      W_g[13,36] := 0.38792211;
      W_g[13,37] := -0.01284714;
      W_g[13,38] := -0.07044123;
      W_g[13,39] := -0.01824626;
      W_g[14,0] := 0.11452243;
      W_g[14,1] := -0.08958103;
      W_g[14,2] := 0.00742450;
      W_g[14,3] := -0.03061342;
      W_g[14,4] := 0.01046369;
      W_g[14,5] := -0.11585659;
      W_g[14,6] := -0.20829633;
      W_g[14,7] := -0.23606929;
      W_g[14,8] := 0.00405464;
      W_g[14,9] := -0.14249870;
      W_g[14,10] := 0.44500434;
      W_g[14,11] := -0.01216610;
      W_g[14,12] := 0.02130103;
      W_g[14,13] := 0.01377995;
      W_g[14,14] := -0.06184130;
      W_g[14,15] := -0.00823075;
      W_g[14,16] := -0.01915279;
      W_g[14,17] := -0.04558576;
      W_g[14,18] := 0.06331799;
      W_g[14,19] := 0.08152927;
      W_g[14,20] := 0.53168559;
      W_g[14,21] := 0.26574171;
      W_g[14,22] := -0.16918069;
      W_g[14,23] := -0.07620575;
      W_g[14,24] := 0.06382546;
      W_g[14,25] := 0.06389488;
      W_g[14,26] := -0.00257182;
      W_g[14,27] := -0.51656342;
      W_g[14,28] := -0.13776320;
      W_g[14,29] := -0.24295253;
      W_g[14,30] := -0.07003054;
      W_g[14,31] := -0.24279301;
      W_g[14,32] := -0.02749909;
      W_g[14,33] := 0.02581101;
      W_g[14,34] := -0.14111596;
      W_g[14,35] := 0.25200224;
      W_g[14,36] := 0.05485417;
      W_g[14,37] := 0.20230512;
      W_g[14,38] := 0.05531698;
      W_g[14,39] := 0.08741502;
      W_g[15,0] := 0.09134059;
      W_g[15,1] := 0.23798586;
      W_g[15,2] := -0.21710049;
      W_g[15,3] := 0.01671123;
      W_g[15,4] := -0.06627945;
      W_g[15,5] := 0.03637264;
      W_g[15,6] := -0.06409252;
      W_g[15,7] := 0.00869699;
      W_g[15,8] := 0.06247383;
      W_g[15,9] := 0.02281686;
      W_g[15,10] := -0.03344842;
      W_g[15,11] := 0.25090969;
      W_g[15,12] := 0.23236279;
      W_g[15,13] := -0.16730684;
      W_g[15,14] := 0.02698623;
      W_g[15,15] := -0.12334466;
      W_g[15,16] := -0.08336571;
      W_g[15,17] := 0.02588012;
      W_g[15,18] := 0.18191151;
      W_g[15,19] := -0.02410393;
      W_g[15,20] := -0.01209911;
      W_g[15,21] := 0.03851634;
      W_g[15,22] := 0.03899917;
      W_g[15,23] := -0.03513279;
      W_g[15,24] := -0.00729930;
      W_g[15,25] := -0.10642073;
      W_g[15,26] := -0.05139272;
      W_g[15,27] := -0.04481147;
      W_g[15,28] := 0.00286298;
      W_g[15,29] := 0.04913988;
      W_g[15,30] := 0.03607814;
      W_g[15,31] := -0.06170525;
      W_g[15,32] := -0.01997224;
      W_g[15,33] := -0.01920844;
      W_g[15,34] := -0.18122375;
      W_g[15,35] := -0.04529240;
      W_g[15,36] := -0.02951458;
      W_g[15,37] := -0.04119204;
      W_g[15,38] := 0.24360354;
      W_g[15,39] := -0.01501589;
      W_g[16,0] := 0.03330758;
      W_g[16,1] := 0.03378529;
      W_g[16,2] := -0.01803414;
      W_g[16,3] := 0.07683524;
      W_g[16,4] := -0.00690420;
      W_g[16,5] := 0.06186575;
      W_g[16,6] := -0.05324589;
      W_g[16,7] := 0.00639146;
      W_g[16,8] := -0.03105667;
      W_g[16,9] := -0.02839811;
      W_g[16,10] := -0.02821902;
      W_g[16,11] := 0.34098804;
      W_g[16,12] := 0.27613014;
      W_g[16,13] := 0.05372236;
      W_g[16,14] := -0.07848245;
      W_g[16,15] := 0.19472931;
      W_g[16,16] := 0.02947051;
      W_g[16,17] := 0.30273750;
      W_g[16,18] := -0.21194892;
      W_g[16,19] := -0.39211345;
      W_g[16,20] := 0.05004872;
      W_g[16,21] := -0.00701097;
      W_g[16,22] := -0.05493126;
      W_g[16,23] := -0.06638756;
      W_g[16,24] := 0.04953207;
      W_g[16,25] := -0.07040619;
      W_g[16,26] := 0.02371565;
      W_g[16,27] := 0.05669258;
      W_g[16,28] := 0.01683023;
      W_g[16,29] := 0.01049871;
      W_g[16,30] := -0.03757136;
      W_g[16,31] := -0.14508742;
      W_g[16,32] := 0.06499721;
      W_g[16,33] := 0.04419298;
      W_g[16,34] := 0.17147748;
      W_g[16,35] := 0.11538684;
      W_g[16,36] := -0.02263807;
      W_g[16,37] := 0.09602714;
      W_g[16,38] := -0.19564001;
      W_g[16,39] := -0.07901151;
      W_g[17,0] := -0.29499203;
      W_g[17,1] := -0.13629365;
      W_g[17,2] := 0.12754540;
      W_g[17,3] := -0.06893644;
      W_g[17,4] := 0.12316505;
      W_g[17,5] := -0.05960383;
      W_g[17,6] := 0.20034896;
      W_g[17,7] := -0.04356226;
      W_g[17,8] := 0.02703761;
      W_g[17,9] := 0.06460494;
      W_g[17,10] := 0.13004684;
      W_g[17,11] := 0.24505885;
      W_g[17,12] := -0.04222988;
      W_g[17,13] := -0.06719559;
      W_g[17,14] := -0.02482782;
      W_g[17,15] := 0.21142994;
      W_g[17,16] := -0.06490519;
      W_g[17,17] := -0.00718676;
      W_g[17,18] := -0.06072595;
      W_g[17,19] := 0.09942021;
      W_g[17,20] := 0.12877691;
      W_g[17,21] := -0.55509835;
      W_g[17,22] := 0.01808993;
      W_g[17,23] := -0.10264266;
      W_g[17,24] := -0.39161390;
      W_g[17,25] := -0.18429647;
      W_g[17,26] := 0.28592888;
      W_g[17,27] := 0.28200120;
      W_g[17,28] := -0.28280002;
      W_g[17,29] := 0.37366402;
      W_g[17,30] := -0.26108804;
      W_g[17,31] := -0.16473882;
      W_g[17,32] := -0.02813312;
      W_g[17,33] := 0.06121552;
      W_g[17,34] := -0.13777223;
      W_g[17,35] := 0.06097139;
      W_g[17,36] := -0.11655490;
      W_g[17,37] := 0.32778808;
      W_g[17,38] := -0.00997418;
      W_g[17,39] := 0.61113542;
      W_g[18,0] := -0.28768328;
      W_g[18,1] := 0.04952108;
      W_g[18,2] := 0.27538794;
      W_g[18,3] := 0.13723339;
      W_g[18,4] := -0.17335135;
      W_g[18,5] := 0.00670465;
      W_g[18,6] := 0.08641540;
      W_g[18,7] := -0.07883801;
      W_g[18,8] := 0.03116638;
      W_g[18,9] := -0.13738742;
      W_g[18,10] := 0.04719661;
      W_g[18,11] := -0.16387163;
      W_g[18,12] := 0.33639768;
      W_g[18,13] := 0.00474426;
      W_g[18,14] := 0.00756510;
      W_g[18,15] := 0.14428972;
      W_g[18,16] := -0.27880877;
      W_g[18,17] := 0.02302493;
      W_g[18,18] := -0.08590068;
      W_g[18,19] := -0.09520416;
      W_g[18,20] := -0.04702628;
      W_g[18,21] := -0.21427108;
      W_g[18,22] := -0.01308084;
      W_g[18,23] := -0.13671976;
      W_g[18,24] := -0.33657643;
      W_g[18,25] := -0.29697937;
      W_g[18,26] := -0.38845918;
      W_g[18,27] := -0.13320677;
      W_g[18,28] := 0.12394036;
      W_g[18,29] := -0.01619850;
      W_g[18,30] := -0.00443483;
      W_g[18,31] := 0.02029626;
      W_g[18,32] := -0.14898181;
      W_g[18,33] := -0.13671023;
      W_g[18,34] := -0.39283904;
      W_g[18,35] := -0.18510637;
      W_g[18,36] := 0.02999584;
      W_g[18,37] := -0.09973078;
      W_g[18,38] := -0.00653579;
      W_g[18,39] := 0.00375571;
      W_g[19,0] := -0.11157153;
      W_g[19,1] := 0.03151476;
      W_g[19,2] := -0.09300674;
      W_g[19,3] := -0.03647256;
      W_g[19,4] := 0.28257591;
      W_g[19,5] := 0.03472368;
      W_g[19,6] := -0.19133006;
      W_g[19,7] := 0.01238337;
      W_g[19,8] := 0.10695083;
      W_g[19,9] := 0.06876826;
      W_g[19,10] := -0.15979454;
      W_g[19,11] := 0.04513165;
      W_g[19,12] := -0.09798693;
      W_g[19,13] := 0.24185713;
      W_g[19,14] := -0.15790631;
      W_g[19,15] := -0.06232450;
      W_g[19,16] := -0.01514155;
      W_g[19,17] := -0.04614652;
      W_g[19,18] := -0.04110415;
      W_g[19,19] := -0.02570745;
      W_g[19,20] := 0.10103595;
      W_g[19,21] := -0.08295028;
      W_g[19,22] := 0.07743288;
      W_g[19,23] := -0.15730743;
      W_g[19,24] := 0.17693761;
      W_g[19,25] := 0.33892640;
      W_g[19,26] := -0.26026049;
      W_g[19,27] := -0.07923400;
      W_g[19,28] := -0.40416408;
      W_g[19,29] := 0.04351845;
      W_g[19,30] := 0.08160401;
      W_g[19,31] := 0.22098459;
      W_g[19,32] := -0.03047447;
      W_g[19,33] := -0.05386001;
      W_g[19,34] := 0.03276813;
      W_g[19,35] := 0.02858822;
      W_g[19,36] := -0.03703291;
      W_g[19,37] := -0.03316212;
      W_g[19,38] := 0.01126183;
      W_g[19,39] := 0.01366358;
      W_g[20,0] := 0.16085938;
      W_g[20,1] := -0.32531878;
      W_g[20,2] := -0.02553925;
      W_g[20,3] := 0.10965997;
      W_g[20,4] := -0.56357527;
      W_g[20,5] := 0.05013693;
      W_g[20,6] := -0.06616703;
      W_g[20,7] := 0.23525825;
      W_g[20,8] := -0.07063977;
      W_g[20,9] := 0.16660647;
      W_g[20,10] := -0.25578102;
      W_g[20,11] := -0.13332653;
      W_g[20,12] := -0.04554458;
      W_g[20,13] := -0.07032327;
      W_g[20,14] := 0.00767713;
      W_g[20,15] := 0.04844571;
      W_g[20,16] := -0.00365021;
      W_g[20,17] := 0.03563506;
      W_g[20,18] := 0.00472104;
      W_g[20,19] := -0.01672288;
      W_g[20,20] := 0.02849239;
      W_g[20,21] := 0.01385569;
      W_g[20,22] := 0.08140633;
      W_g[20,23] := -0.12280270;
      W_g[20,24] := -0.13321750;
      W_g[20,25] := -0.07573776;
      W_g[20,26] := -0.11991729;
      W_g[20,27] := 0.08519396;
      W_g[20,28] := -0.22153257;
      W_g[20,29] := 0.06635125;
      W_g[20,30] := 0.03284018;
      W_g[20,31] := -0.04984721;
      W_g[20,32] := -0.02468482;
      W_g[20,33] := -0.03918115;
      W_g[20,34] := -0.33116385;
      W_g[20,35] := -0.07214631;
      W_g[20,36] := -0.11911645;
      W_g[20,37] := 0.02867687;
      W_g[20,38] := 0.10832489;
      W_g[20,39] := -0.03266538;
      W_g[21,0] := -0.12645213;
      W_g[21,1] := 0.08150304;
      W_g[21,2] := 0.02647559;
      W_g[21,3] := 0.08127797;
      W_g[21,4] := 0.04152407;
      W_g[21,5] := -0.00439330;
      W_g[21,6] := -0.06754721;
      W_g[21,7] := -0.01934627;
      W_g[21,8] := 0.02639229;
      W_g[21,9] := -0.05531998;
      W_g[21,10] := -0.02184705;
      W_g[21,11] := 0.05361381;
      W_g[21,12] := -0.08168689;
      W_g[21,13] := 0.04307065;
      W_g[21,14] := 0.34190872;
      W_g[21,15] := 0.01199497;
      W_g[21,16] := 0.02785254;
      W_g[21,17] := -0.01922297;
      W_g[21,18] := 0.00887910;
      W_g[21,19] := -0.63622159;
      W_g[21,20] := 0.10488117;
      W_g[21,21] := 0.21346407;
      W_g[21,22] := -0.01027352;
      W_g[21,23] := 0.02464858;
      W_g[21,24] := -0.16255559;
      W_g[21,25] := -0.44461492;
      W_g[21,26] := 0.04926345;
      W_g[21,27] := -0.12672877;
      W_g[21,28] := 0.04893465;
      W_g[21,29] := -0.02553335;
      W_g[21,30] := 0.02661697;
      W_g[21,31] := -0.02238514;
      W_g[21,32] := -0.01370737;
      W_g[21,33] := -0.02438860;
      W_g[21,34] := -0.03352462;
      W_g[21,35] := -0.00976400;
      W_g[21,36] := -0.00314182;
      W_g[21,37] := -0.01966831;
      W_g[21,38] := 0.08250269;
      W_g[21,39] := 0.03922363;
      W_g[22,0] := 0.21398924;
      W_g[22,1] := -0.01974818;
      W_g[22,2] := 0.04753013;
      W_g[22,3] := -0.24118032;
      W_g[22,4] := 0.14757568;
      W_g[22,5] := 0.11998211;
      W_g[22,6] := -0.20516486;
      W_g[22,7] := -0.00517598;
      W_g[22,8] := -0.17191212;
      W_g[22,9] := 0.02895894;
      W_g[22,10] := 0.06158756;
      W_g[22,11] := 0.22470629;
      W_g[22,12] := -0.01264452;
      W_g[22,13] := -0.01041790;
      W_g[22,14] := 0.00696788;
      W_g[22,15] := 0.01863093;
      W_g[22,16] := -0.17598189;
      W_g[22,17] := -0.01077684;
      W_g[22,18] := 0.00929625;
      W_g[22,19] := -0.06654035;
      W_g[22,20] := 0.04213786;
      W_g[22,21] := 0.16789195;
      W_g[22,22] := 0.16808763;
      W_g[22,23] := 0.09369668;
      W_g[22,24] := 0.33967805;
      W_g[22,25] := 0.04618895;
      W_g[22,26] := 0.17455877;
      W_g[22,27] := 0.09184463;
      W_g[22,28] := 0.00975296;
      W_g[22,29] := 0.09664790;
      W_g[22,30] := 0.16180007;
      W_g[22,31] := -0.15128982;
      W_g[22,32] := -0.13754758;
      W_g[22,33] := -0.14797860;
      W_g[22,34] := 0.29874405;
      W_g[22,35] := -0.17532231;
      W_g[22,36] := -0.05865765;
      W_g[22,37] := -0.28989062;
      W_g[22,38] := -0.06785104;
      W_g[22,39] := 0.19310509;
      W_g[23,0] := 0.02262829;
      W_g[23,1] := -0.14467132;
      W_g[23,2] := 0.15171790;
      W_g[23,3] := -0.05470154;
      W_g[23,4] := 0.11472824;
      W_g[23,5] := 0.02458709;
      W_g[23,6] := 0.00195381;
      W_g[23,7] := -0.03838236;
      W_g[23,8] := -0.08246408;
      W_g[23,9] := -0.03637726;
      W_g[23,10] := 0.05126188;
      W_g[23,11] := 0.08157095;
      W_g[23,12] := 0.17084308;
      W_g[23,13] := 0.04612783;
      W_g[23,14] := 0.00166863;
      W_g[23,15] := -0.11824610;
      W_g[23,16] := 0.25113744;
      W_g[23,17] := -0.00895557;
      W_g[23,18] := -0.09017404;
      W_g[23,19] := -0.00864124;
      W_g[23,20] := -0.17411692;
      W_g[23,21] := -0.23732638;
      W_g[23,22] := -0.01919251;
      W_g[23,23] := 0.05404213;
      W_g[23,24] := -0.23653357;
      W_g[23,25] := -0.05463766;
      W_g[23,26] := -0.09652406;
      W_g[23,27] := 0.06527363;
      W_g[23,28] := -0.11678946;
      W_g[23,29] := 0.04067237;
      W_g[23,30] := -0.04251467;
      W_g[23,31] := -0.02616764;
      W_g[23,32] := -0.04019048;
      W_g[23,33] := -0.09613159;
      W_g[23,34] := -0.13061938;
      W_g[23,35] := -0.00608878;
      W_g[23,36] := -0.00901942;
      W_g[23,37] := -0.03102667;
      W_g[23,38] := 0.06219607;
      W_g[23,39] := -0.03399585;
      W_g[24,0] := -0.07987209;
      W_g[24,1] := 0.14030914;
      W_g[24,2] := -0.00618952;
      W_g[24,3] := -0.03472964;
      W_g[24,4] := -0.25152627;
      W_g[24,5] := 0.02353315;
      W_g[24,6] := 0.27113226;
      W_g[24,7] := -0.09270474;
      W_g[24,8] := 0.09813852;
      W_g[24,9] := -0.03003301;
      W_g[24,10] := 0.14422308;
      W_g[24,11] := 0.12668727;
      W_g[24,12] := 0.06848053;
      W_g[24,13] := -0.05021099;
      W_g[24,14] := 0.00261446;
      W_g[24,15] := -0.14804363;
      W_g[24,16] := 0.09895858;
      W_g[24,17] := -0.01510628;
      W_g[24,18] := -0.00454297;
      W_g[24,19] := -0.09103126;
      W_g[24,20] := 0.00004775;
      W_g[24,21] := 0.05401549;
      W_g[24,22] := 0.05428678;
      W_g[24,23] := 0.10576063;
      W_g[24,24] := 0.19301949;
      W_g[24,25] := 0.09099979;
      W_g[24,26] := 0.15261312;
      W_g[24,27] := -0.20747845;
      W_g[24,28] := -0.37421781;
      W_g[24,29] := -0.01107945;
      W_g[24,30] := 0.10706456;
      W_g[24,31] := 0.19086725;
      W_g[24,32] := -0.02514360;
      W_g[24,33] := -0.01640238;
      W_g[24,34] := 0.08067109;
      W_g[24,35] := -0.06559525;
      W_g[24,36] := -0.08709598;
      W_g[24,37] := -0.15054889;
      W_g[24,38] := -0.25885892;
      W_g[24,39] := 0.01723043;
      W_g[25,0] := 0.06067028;
      W_g[25,1] := 0.15727347;
      W_g[25,2] := 0.06245382;
      W_g[25,3] := 0.04814018;
      W_g[25,4] := -0.05496313;
      W_g[25,5] := 0.02508350;
      W_g[25,6] := -0.11731715;
      W_g[25,7] := 0.11065199;
      W_g[25,8] := -0.06903063;
      W_g[25,9] := 0.04847066;
      W_g[25,10] := -0.23851803;
      W_g[25,11] := -0.11894847;
      W_g[25,12] := -0.00354003;
      W_g[25,13] := -0.23670243;
      W_g[25,14] := -0.11929761;
      W_g[25,15] := 0.06615548;
      W_g[25,16] := 0.02567591;
      W_g[25,17] := -0.11101572;
      W_g[25,18] := 0.02320875;
      W_g[25,19] := -0.00523274;
      W_g[25,20] := 0.17951657;
      W_g[25,21] := -0.23383175;
      W_g[25,22] := -0.04463376;
      W_g[25,23] := 0.07589541;
      W_g[25,24] := -0.38295865;
      W_g[25,25] := -0.26238292;
      W_g[25,26] := -0.11914421;
      W_g[25,27] := 0.12171790;
      W_g[25,28] := 0.01532443;
      W_g[25,29] := -0.13715334;
      W_g[25,30] := -0.07302305;
      W_g[25,31] := -0.10361797;
      W_g[25,32] := -0.04133119;
      W_g[25,33] := 0.07758912;
      W_g[25,34] := 0.13717994;
      W_g[25,35] := -0.18056835;
      W_g[25,36] := -0.22574168;
      W_g[25,37] := -0.02318463;
      W_g[25,38] := -0.03606231;
      W_g[25,39] := 0.01114746;
      W_g[26,0] := 0.04868018;
      W_g[26,1] := 0.10704073;
      W_g[26,2] := -0.09924373;
      W_g[26,3] := 0.01612309;
      W_g[26,4] := -0.28056058;
      W_g[26,5] := 0.00307460;
      W_g[26,6] := 0.13066944;
      W_g[26,7] := 0.08240058;
      W_g[26,8] := -0.01877597;
      W_g[26,9] := 0.07625350;
      W_g[26,10] := -0.01633129;
      W_g[26,11] := -0.06490228;
      W_g[26,12] := 0.00356371;
      W_g[26,13] := 0.60836279;
      W_g[26,14] := -0.00784845;
      W_g[26,15] := 0.14515170;
      W_g[26,16] := 0.00666268;
      W_g[26,17] := -0.08984287;
      W_g[26,18] := -0.10734571;
      W_g[26,19] := 0.06982262;
      W_g[26,20] := -0.15198155;
      W_g[26,21] := 0.08035437;
      W_g[26,22] := -0.00864624;
      W_g[26,23] := 0.17810401;
      W_g[26,24] := 0.32582802;
      W_g[26,25] := 0.04504528;
      W_g[26,26] := -0.08173288;
      W_g[26,27] := 0.00872430;
      W_g[26,28] := -0.05935643;
      W_g[26,29] := 0.00892613;
      W_g[26,30] := -0.01252034;
      W_g[26,31] := -0.20071557;
      W_g[26,32] := -0.01037293;
      W_g[26,33] := 0.02427795;
      W_g[26,34] := 0.02944206;
      W_g[26,35] := -0.13762893;
      W_g[26,36] := 0.01954584;
      W_g[26,37] := 0.01543705;
      W_g[26,38] := 0.13130702;
      W_g[26,39] := -0.00475240;
      W_g[27,0] := 0.26684397;
      W_g[27,1] := -0.10793137;
      W_g[27,2] := -0.33427569;
      W_g[27,3] := 0.16579777;
      W_g[27,4] := 0.08486222;
      W_g[27,5] := -0.08615804;
      W_g[27,6] := -0.04872312;
      W_g[27,7] := -0.09806403;
      W_g[27,8] := 0.11429329;
      W_g[27,9] := -0.15268981;
      W_g[27,10] := 0.14884192;
      W_g[27,11] := -0.19054756;
      W_g[27,12] := 0.11245804;
      W_g[27,13] := 0.11537316;
      W_g[27,14] := 0.00333165;
      W_g[27,15] := 0.11125144;
      W_g[27,16] := 0.11089247;
      W_g[27,17] := 0.00310823;
      W_g[27,18] := 0.30689535;
      W_g[27,19] := -0.03992568;
      W_g[27,20] := 0.04893808;
      W_g[27,21] := -0.12398542;
      W_g[27,22] := -0.07112632;
      W_g[27,23] := 0.11366460;
      W_g[27,24] := -0.41621515;
      W_g[27,25] := -0.24068177;
      W_g[27,26] := -0.17630154;
      W_g[27,27] := 0.18514685;
      W_g[27,28] := 0.07259171;
      W_g[27,29] := 0.06956388;
      W_g[27,30] := -0.09684508;
      W_g[27,31] := 0.14715137;
      W_g[27,32] := -0.04076103;
      W_g[27,33] := -0.04563152;
      W_g[27,34] := -0.37191504;
      W_g[27,35] := 0.01961966;
      W_g[27,36] := -0.03775807;
      W_g[27,37] := 0.11485546;
      W_g[27,38] := -0.25651574;
      W_g[27,39] := -0.01313073;
      W_g[28,0] := -0.13160358;
      W_g[28,1] := 0.07208443;
      W_g[28,2] := -0.19002992;
      W_g[28,3] := -0.01230462;
      W_g[28,4] := -0.19478217;
      W_g[28,5] := 0.72986090;
      W_g[28,6] := -0.41573420;
      W_g[28,7] := -0.00614311;
      W_g[28,8] := 0.21563159;
      W_g[28,9] := 0.06237340;
      W_g[28,10] := 0.34260488;
      W_g[28,11] := -0.08146781;
      W_g[28,12] := -0.29444560;
      W_g[28,13] := -0.02234161;
      W_g[28,14] := 0.00739318;
      W_g[28,15] := 0.03697482;
      W_g[28,16] := 0.07958936;
      W_g[28,17] := 0.03669633;
      W_g[28,18] := -0.04358352;
      W_g[28,19] := 0.07740789;
      W_g[28,20] := -0.38667741;
      W_g[28,21] := -0.05676787;
      W_g[28,22] := 0.01061609;
      W_g[28,23] := -0.03819450;
      W_g[28,24] := -0.02419050;
      W_g[28,25] := -0.19251022;
      W_g[28,26] := -0.01905529;
      W_g[28,27] := 0.21895112;
      W_g[28,28] := 0.00464667;
      W_g[28,29] := -0.09290081;
      W_g[28,30] := -0.08549001;
      W_g[28,31] := 0.05558621;
      W_g[28,32] := -0.05720450;
      W_g[28,33] := -0.00354341;
      W_g[28,34] := 0.01472593;
      W_g[28,35] := 0.01051784;
      W_g[28,36] := -0.04851991;
      W_g[28,37] := 0.06329209;
      W_g[28,38] := 0.03593949;
      W_g[28,39] := 0.03454753;
      W_g[29,0] := -0.05209588;
      W_g[29,1] := 0.17165838;
      W_g[29,2] := 0.35414502;
      W_g[29,3] := 0.23215105;
      W_g[29,4] := 0.35465872;
      W_g[29,5] := 0.04213377;
      W_g[29,6] := 0.17051828;
      W_g[29,7] := 0.44905955;
      W_g[29,8] := -0.18509297;
      W_g[29,9] := 0.34960920;
      W_g[29,10] := 0.06534662;
      W_g[29,11] := 0.00280209;
      W_g[29,12] := 0.07823030;
      W_g[29,13] := -0.04565757;
      W_g[29,14] := 0.00520064;
      W_g[29,15] := 0.03880082;
      W_g[29,16] := -0.02205570;
      W_g[29,17] := 0.03516322;
      W_g[29,18] := 0.40971720;
      W_g[29,19] := -0.02489867;
      W_g[29,20] := -0.11450347;
      W_g[29,21] := 0.14212352;
      W_g[29,22] := -0.04341381;
      W_g[29,23] := 0.04860599;
      W_g[29,24] := 0.03678778;
      W_g[29,25] := 0.00164296;
      W_g[29,26] := 0.13215743;
      W_g[29,27] := -0.07260210;
      W_g[29,28] := -0.34370157;
      W_g[29,29] := -0.30255622;
      W_g[29,30] := -0.00881223;
      W_g[29,31] := -0.05561844;
      W_g[29,32] := -0.05011707;
      W_g[29,33] := -0.05156367;
      W_g[29,34] := -0.06613368;
      W_g[29,35] := 0.12263016;
      W_g[29,36] := -0.00414138;
      W_g[29,37] := -0.02915506;
      W_g[29,38] := -0.02212529;
      W_g[29,39] := 0.12280423;
      W_g[30,0] := -0.07765778;
      W_g[30,1] := -0.01351530;
      W_g[30,2] := 0.06473100;
      W_g[30,3] := 0.04457490;
      W_g[30,4] := -0.04750980;
      W_g[30,5] := -0.06268556;
      W_g[30,6] := -0.10883031;
      W_g[30,7] := -0.07578032;
      W_g[30,8] := 0.06264021;
      W_g[30,9] := -0.07505340;
      W_g[30,10] := 0.02022277;
      W_g[30,11] := 0.00762805;
      W_g[30,12] := 0.10820425;
      W_g[30,13] := -0.00375025;
      W_g[30,14] := 0.00127143;
      W_g[30,15] := 0.26273328;
      W_g[30,16] := 0.14333837;
      W_g[30,17] := -0.06559381;
      W_g[30,18] := 0.00541820;
      W_g[30,19] := 0.04841781;
      W_g[30,20] := -0.13715798;
      W_g[30,21] := 0.10902844;
      W_g[30,22] := 0.07313410;
      W_g[30,23] := -0.18172082;
      W_g[30,24] := 0.33205184;
      W_g[30,25] := 0.33727106;
      W_g[30,26] := 0.18524152;
      W_g[30,27] := 0.00587510;
      W_g[30,28] := 0.01138745;
      W_g[30,29] := -0.00862603;
      W_g[30,30] := 0.03883495;
      W_g[30,31] := 0.01710799;
      W_g[30,32] := -0.01818751;
      W_g[30,33] := -0.00650796;
      W_g[30,34] := 0.09579980;
      W_g[30,35] := -0.09178187;
      W_g[30,36] := 0.02701038;
      W_g[30,37] := -0.05651341;
      W_g[30,38] := 0.02332304;
      W_g[30,39] := 0.00988352;
      W_g[31,0] := -0.07066347;
      W_g[31,1] := -0.25243866;
      W_g[31,2] := -0.15006079;
      W_g[31,3] := -0.06871642;
      W_g[31,4] := 0.02799054;
      W_g[31,5] := -0.18761340;
      W_g[31,6] := 0.20777020;
      W_g[31,7] := -0.01511925;
      W_g[31,8] := 0.24296197;
      W_g[31,9] := 0.17157343;
      W_g[31,10] := 0.34240860;
      W_g[31,11] := 0.17374654;
      W_g[31,12] := 0.01123912;
      W_g[31,13] := 0.05064730;
      W_g[31,14] := -0.11290316;
      W_g[31,15] := -0.07592911;
      W_g[31,16] := -0.05080255;
      W_g[31,17] := -0.03835510;
      W_g[31,18] := -0.10784303;
      W_g[31,19] := -0.14260224;
      W_g[31,20] := 0.01680487;
      W_g[31,21] := -0.12900466;
      W_g[31,22] := 0.15861642;
      W_g[31,23] := -0.03345355;
      W_g[31,24] := 0.03338373;
      W_g[31,25] := 0.33927539;
      W_g[31,26] := -0.03024811;
      W_g[31,27] := 0.21193095;
      W_g[31,28] := 0.14089774;
      W_g[31,29] := -0.04104134;
      W_g[31,30] := 0.13590372;
      W_g[31,31] := 0.00341222;
      W_g[31,32] := -0.06720376;
      W_g[31,33] := -0.06392696;
      W_g[31,34] := 0.32630247;
      W_g[31,35] := -0.29304048;
      W_g[31,36] := -0.08099687;
      W_g[31,37] := -0.18760577;
      W_g[31,38] := 0.05159000;
      W_g[31,39] := 0.03953602;
      W_o[0,0] := 0.36960590;
      W_o[0,1] := -0.20815031;
      W_o[0,2] := 0.02135882;
      W_o[0,3] := -0.40729395;
      W_o[0,4] := -0.08193119;
      W_o[0,5] := -0.05334249;
      W_o[0,6] := 0.31897318;
      W_o[0,7] := -0.30747417;
      W_o[0,8] := 0.11512720;
      W_o[0,9] := -0.38517836;
      W_o[0,10] := -0.11075519;
      W_o[0,11] := 0.21201350;
      W_o[0,12] := 0.02026256;
      W_o[0,13] := -0.24249811;
      W_o[0,14] := -0.30325094;
      W_o[0,15] := 0.01195520;
      W_o[0,16] := 0.01862234;
      W_o[0,17] := -0.19610310;
      W_o[0,18] := 0.01511792;
      W_o[0,19] := 0.10368652;
      W_o[0,20] := 0.16080864;
      W_o[0,21] := 0.60025555;
      W_o[0,22] := 0.04030931;
      W_o[0,23] := -0.12621889;
      W_o[0,24] := -0.32480696;
      W_o[0,25] := -0.17387474;
      W_o[0,26] := -0.37594935;
      W_o[0,27] := 0.24470490;
      W_o[0,28] := 0.20932631;
      W_o[0,29] := -0.28829920;
      W_o[0,30] := -0.18935557;
      W_o[0,31] := -0.13508852;
      W_o[0,32] := -0.09435762;
      W_o[0,33] := 0.41882566;
      W_o[0,34] := 0.12677918;
      W_o[0,35] := -0.09689110;
      W_o[0,36] := 0.00309573;
      W_o[0,37] := 0.02559190;
      W_o[0,38] := -0.03516277;
      W_o[0,39] := 0.36212319;
      W_o[1,0] := 0.00818965;
      W_o[1,1] := -0.05766975;
      W_o[1,2] := -0.25532568;
      W_o[1,3] := 0.00466345;
      W_o[1,4] := -0.64983314;
      W_o[1,5] := 0.67811555;
      W_o[1,6] := -0.07523961;
      W_o[1,7] := 0.05286549;
      W_o[1,8] := -0.08405841;
      W_o[1,9] := -0.13089836;
      W_o[1,10] := 0.05647256;
      W_o[1,11] := -0.41155520;
      W_o[1,12] := -0.28863174;
      W_o[1,13] := 0.05577922;
      W_o[1,14] := 0.05531852;
      W_o[1,15] := -0.50346696;
      W_o[1,16] := -0.12134568;
      W_o[1,17] := -0.32418999;
      W_o[1,18] := -0.17313546;
      W_o[1,19] := -0.11050858;
      W_o[1,20] := -0.10319410;
      W_o[1,21] := 0.02116561;
      W_o[1,22] := -0.04030692;
      W_o[1,23] := -0.05150330;
      W_o[1,24] := -0.31542593;
      W_o[1,25] := -0.09472059;
      W_o[1,26] := -0.25657916;
      W_o[1,27] := 0.33742470;
      W_o[1,28] := 0.46666449;
      W_o[1,29] := -0.24623868;
      W_o[1,30] := 0.10010793;
      W_o[1,31] := 0.11690982;
      W_o[1,32] := 0.05103257;
      W_o[1,33] := 0.04395993;
      W_o[1,34] := 0.05502438;
      W_o[1,35] := -0.04573586;
      W_o[1,36] := 0.07247765;
      W_o[1,37] := -0.12633540;
      W_o[1,38] := -0.02435859;
      W_o[1,39] := -0.19470915;
      W_o[2,0] := 0.56892127;
      W_o[2,1] := 0.21849076;
      W_o[2,2] := -0.51244366;
      W_o[2,3] := 0.12966341;
      W_o[2,4] := -0.37199587;
      W_o[2,5] := 0.31576705;
      W_o[2,6] := 0.47295788;
      W_o[2,7] := -0.11773749;
      W_o[2,8] := 0.03722378;
      W_o[2,9] := -0.06956325;
      W_o[2,10] := 0.08040347;
      W_o[2,11] := -0.17961407;
      W_o[2,12] := -0.10757016;
      W_o[2,13] := 0.15337250;
      W_o[2,14] := 0.13618986;
      W_o[2,15] := 0.22858761;
      W_o[2,16] := -0.00072664;
      W_o[2,17] := 0.11959419;
      W_o[2,18] := 0.14819941;
      W_o[2,19] := -0.17484270;
      W_o[2,20] := -0.60648781;
      W_o[2,21] := 0.80117035;
      W_o[2,22] := 0.26442236;
      W_o[2,23] := -0.26784527;
      W_o[2,24] := 1.16267180;
      W_o[2,25] := 1.05618489;
      W_o[2,26] := -0.05316524;
      W_o[2,27] := 0.29363456;
      W_o[2,28] := 0.18678209;
      W_o[2,29] := -0.03277919;
      W_o[2,30] := 0.24237865;
      W_o[2,31] := -0.15350257;
      W_o[2,32] := 0.08219703;
      W_o[2,33] := 0.09145115;
      W_o[2,34] := 0.90349656;
      W_o[2,35] := 0.33768374;
      W_o[2,36] := 0.46036184;
      W_o[2,37] := 0.33086196;
      W_o[2,38] := 0.00527997;
      W_o[2,39] := 0.38400045;
      W_o[3,0] := -0.13949616;
      W_o[3,1] := -0.00636318;
      W_o[3,2] := -0.10001112;
      W_o[3,3] := -0.33833316;
      W_o[3,4] := 0.12226738;
      W_o[3,5] := -0.00821515;
      W_o[3,6] := 0.12485677;
      W_o[3,7] := -0.03404867;
      W_o[3,8] := 0.19117068;
      W_o[3,9] := 0.17734979;
      W_o[3,10] := 0.15269712;
      W_o[3,11] := 0.11457094;
      W_o[3,12] := -0.54962271;
      W_o[3,13] := -0.15097325;
      W_o[3,14] := -0.06021854;
      W_o[3,15] := 0.31263557;
      W_o[3,16] := 0.21840449;
      W_o[3,17] := 0.18637469;
      W_o[3,18] := 0.00558414;
      W_o[3,19] := 0.03386161;
      W_o[3,20] := -0.00529720;
      W_o[3,21] := 0.50283587;
      W_o[3,22] := 0.23464191;
      W_o[3,23] := 0.22633280;
      W_o[3,24] := -0.34072113;
      W_o[3,25] := -0.20596467;
      W_o[3,26] := 0.03239496;
      W_o[3,27] := -0.27217436;
      W_o[3,28] := -0.06646252;
      W_o[3,29] := 0.11120258;
      W_o[3,30] := 0.19604938;
      W_o[3,31] := -0.76824152;
      W_o[3,32] := -0.11828657;
      W_o[3,33] := -0.19211680;
      W_o[3,34] := -0.04434033;
      W_o[3,35] := -0.15079519;
      W_o[3,36] := 0.05358901;
      W_o[3,37] := -0.20020793;
      W_o[3,38] := 0.00906296;
      W_o[3,39] := 0.94856155;
      W_o[4,0] := 0.07946882;
      W_o[4,1] := -0.02597320;
      W_o[4,2] := 0.12188822;
      W_o[4,3] := -0.23110408;
      W_o[4,4] := -0.04543841;
      W_o[4,5] := -0.08577575;
      W_o[4,6] := 0.18635339;
      W_o[4,7] := 0.19728531;
      W_o[4,8] := -0.16972877;
      W_o[4,9] := 0.41852465;
      W_o[4,10] := -0.34732747;
      W_o[4,11] := 0.06388048;
      W_o[4,12] := -0.15282933;
      W_o[4,13] := -0.08337624;
      W_o[4,14] := 0.03326624;
      W_o[4,15] := 0.27675766;
      W_o[4,16] := 0.02420580;
      W_o[4,17] := 0.05359625;
      W_o[4,18] := 0.15546103;
      W_o[4,19] := -0.05985435;
      W_o[4,20] := 0.14620510;
      W_o[4,21] := -0.17060445;
      W_o[4,22] := 0.22486657;
      W_o[4,23] := 0.06779833;
      W_o[4,24] := -0.02401932;
      W_o[4,25] := 0.27871072;
      W_o[4,26] := -0.39190814;
      W_o[4,27] := 0.10446193;
      W_o[4,28] := 0.03558551;
      W_o[4,29] := -0.18836324;
      W_o[4,30] := -0.27463332;
      W_o[4,31] := 0.51233327;
      W_o[4,32] := -0.62388706;
      W_o[4,33] := -0.34844089;
      W_o[4,34] := -0.32486844;
      W_o[4,35] := -0.13829319;
      W_o[4,36] := 0.09612888;
      W_o[4,37] := -0.25610924;
      W_o[4,38] := 0.17635575;
      W_o[4,39] := -0.03314881;
      W_o[5,0] := 0.29998592;
      W_o[5,1] := 0.62471324;
      W_o[5,2] := -0.35768643;
      W_o[5,3] := 0.05470141;
      W_o[5,4] := -0.06384566;
      W_o[5,5] := 0.08787517;
      W_o[5,6] := 0.16561310;
      W_o[5,7] := 0.24364167;
      W_o[5,8] := -0.16042867;
      W_o[5,9] := -0.04153518;
      W_o[5,10] := -0.04475499;
      W_o[5,11] := -0.00533060;
      W_o[5,12] := -0.17453381;
      W_o[5,13] := -0.32039422;
      W_o[5,14] := 0.28441662;
      W_o[5,15] := -0.11029031;
      W_o[5,16] := -0.02602161;
      W_o[5,17] := 0.30602705;
      W_o[5,18] := -0.00562938;
      W_o[5,19] := -0.02381407;
      W_o[5,20] := -0.56547868;
      W_o[5,21] := 0.07034699;
      W_o[5,22] := 0.13362850;
      W_o[5,23] := 0.29412499;
      W_o[5,24] := 1.33312082;
      W_o[5,25] := 0.36348087;
      W_o[5,26] := -0.25760710;
      W_o[5,27] := 0.22991443;
      W_o[5,28] := 0.37971079;
      W_o[5,29] := -0.19349299;
      W_o[5,30] := 0.03992765;
      W_o[5,31] := -0.07852311;
      W_o[5,32] := -0.07730967;
      W_o[5,33] := -0.05783857;
      W_o[5,34] := 0.21159130;
      W_o[5,35] := 0.09816961;
      W_o[5,36] := 0.33947071;
      W_o[5,37] := 0.03416896;
      W_o[5,38] := -0.13325274;
      W_o[5,39] := -0.39347383;
      W_o[6,0] := 0.04164087;
      W_o[6,1] := -0.02401152;
      W_o[6,2] := -0.03398127;
      W_o[6,3] := 0.05101350;
      W_o[6,4] := 0.07298061;
      W_o[6,5] := 0.09403470;
      W_o[6,6] := 0.36079749;
      W_o[6,7] := -0.04026723;
      W_o[6,8] := -0.00128813;
      W_o[6,9] := 0.16855729;
      W_o[6,10] := -0.12973289;
      W_o[6,11] := -0.31573737;
      W_o[6,12] := -0.06414645;
      W_o[6,13] := -0.01722028;
      W_o[6,14] := 0.01204535;
      W_o[6,15] := 0.08021659;
      W_o[6,16] := -0.01998950;
      W_o[6,17] := -0.01548403;
      W_o[6,18] := 0.30389985;
      W_o[6,19] := 0.00609801;
      W_o[6,20] := -1.08852530;
      W_o[6,21] := -0.00168008;
      W_o[6,22] := 0.08513393;
      W_o[6,23] := -0.07552507;
      W_o[6,24] := 0.67528367;
      W_o[6,25] := 0.55059099;
      W_o[6,26] := -0.13680276;
      W_o[6,27] := 0.12081103;
      W_o[6,28] := 0.13821204;
      W_o[6,29] := -0.29566112;
      W_o[6,30] := 0.17353611;
      W_o[6,31] := 0.11022282;
      W_o[6,32] := 0.20766126;
      W_o[6,33] := 0.16963202;
      W_o[6,34] := 0.83168727;
      W_o[6,35] := 0.39787611;
      W_o[6,36] := 0.03474040;
      W_o[6,37] := 0.40801755;
      W_o[6,38] := -0.11616077;
      W_o[6,39] := 0.73190320;
      W_o[7,0] := -1.03722596;
      W_o[7,1] := -0.76202756;
      W_o[7,2] := -0.60125434;
      W_o[7,3] := 0.08797976;
      W_o[7,4] := -0.19053090;
      W_o[7,5] := 0.10532437;
      W_o[7,6] := -0.42051023;
      W_o[7,7] := -0.07490456;
      W_o[7,8] := -0.62126988;
      W_o[7,9] := 0.19605152;
      W_o[7,10] := 0.11288203;
      W_o[7,11] := 0.02348748;
      W_o[7,12] := 0.25075635;
      W_o[7,13] := -0.10330101;
      W_o[7,14] := 0.11590070;
      W_o[7,15] := -0.09985835;
      W_o[7,16] := 0.00186775;
      W_o[7,17] := -0.29451331;
      W_o[7,18] := 0.46819898;
      W_o[7,19] := -0.22970740;
      W_o[7,20] := -0.06142933;
      W_o[7,21] := 0.20279525;
      W_o[7,22] := 0.23697145;
      W_o[7,23] := -0.05793158;
      W_o[7,24] := -0.12877418;
      W_o[7,25] := -0.17714323;
      W_o[7,26] := 0.09780758;
      W_o[7,27] := 0.51964223;
      W_o[7,28] := 0.51194477;
      W_o[7,29] := 0.16508958;
      W_o[7,30] := 0.20431308;
      W_o[7,31] := 0.00562293;
      W_o[7,32] := 0.00411460;
      W_o[7,33] := 0.08410010;
      W_o[7,34] := 0.15867023;
      W_o[7,35] := 0.08692707;
      W_o[7,36] := -0.13108705;
      W_o[7,37] := 0.01137071;
      W_o[7,38] := 0.12501325;
      W_o[7,39] := 0.25273043;
      W_o[8,0] := 0.01043700;
      W_o[8,1] := -0.02130833;
      W_o[8,2] := 0.38301000;
      W_o[8,3] := -0.37692562;
      W_o[8,4] := 0.16604906;
      W_o[8,5] := 0.05526777;
      W_o[8,6] := -0.09484355;
      W_o[8,7] := -0.15874933;
      W_o[8,8] := -0.15982778;
      W_o[8,9] := -0.30258146;
      W_o[8,10] := -0.19271901;
      W_o[8,11] := -0.12934390;
      W_o[8,12] := -0.19251528;
      W_o[8,13] := 0.18497486;
      W_o[8,14] := -0.12623328;
      W_o[8,15] := 0.16649424;
      W_o[8,16] := 0.45124924;
      W_o[8,17] := 0.08460020;
      W_o[8,18] := 0.33701915;
      W_o[8,19] := -0.14333396;
      W_o[8,20] := -0.19551557;
      W_o[8,21] := 0.05818683;
      W_o[8,22] := 0.33913088;
      W_o[8,23] := -0.16286211;
      W_o[8,24] := 0.96390134;
      W_o[8,25] := 1.18908966;
      W_o[8,26] := -0.09017515;
      W_o[8,27] := 0.02218129;
      W_o[8,28] := -0.07352100;
      W_o[8,29] := -0.15695611;
      W_o[8,30] := 0.32942769;
      W_o[8,31] := 0.10831923;
      W_o[8,32] := 0.21786334;
      W_o[8,33] := 0.03463054;
      W_o[8,34] := 1.36861372;
      W_o[8,35] := 0.36430228;
      W_o[8,36] := 0.24335380;
      W_o[8,37] := 0.26164109;
      W_o[8,38] := -0.18121149;
      W_o[8,39] := 0.02990196;
      W_o[9,0] := -1.04737031;
      W_o[9,1] := -0.20712732;
      W_o[9,2] := -0.95441955;
      W_o[9,3] := 0.01938875;
      W_o[9,4] := -0.11212977;
      W_o[9,5] := -0.06146387;
      W_o[9,6] := 0.30708382;
      W_o[9,7] := 0.22604913;
      W_o[9,8] := -1.80963576;
      W_o[9,9] := 0.22610889;
      W_o[9,10] := -0.35715115;
      W_o[9,11] := -0.23053938;
      W_o[9,12] := -0.23544851;
      W_o[9,13] := 0.16765821;
      W_o[9,14] := 0.18199258;
      W_o[9,15] := -0.12609567;
      W_o[9,16] := 0.19273403;
      W_o[9,17] := 0.70470548;
      W_o[9,18] := 0.40443879;
      W_o[9,19] := -0.29892516;
      W_o[9,20] := -0.23205499;
      W_o[9,21] := 0.01917006;
      W_o[9,22] := 0.04775739;
      W_o[9,23] := 0.22877300;
      W_o[9,24] := 0.22836986;
      W_o[9,25] := 0.10442287;
      W_o[9,26] := 0.04376736;
      W_o[9,27] := 0.19467911;
      W_o[9,28] := 0.00064683;
      W_o[9,29] := -0.15721194;
      W_o[9,30] := 0.12573351;
      W_o[9,31] := -0.09639835;
      W_o[9,32] := 0.03846860;
      W_o[9,33] := -0.10591342;
      W_o[9,34] := -0.06322171;
      W_o[9,35] := 0.07575873;
      W_o[9,36] := 0.01897552;
      W_o[9,37] := -0.05338341;
      W_o[9,38] := -0.12568939;
      W_o[9,39] := 0.04643562;
      W_o[10,0] := 0.15450947;
      W_o[10,1] := 0.03275542;
      W_o[10,2] := -0.09800130;
      W_o[10,3] := 0.26718503;
      W_o[10,4] := 0.10269620;
      W_o[10,5] := -0.05641613;
      W_o[10,6] := 0.24852888;
      W_o[10,7] := -0.19179238;
      W_o[10,8] := 0.01932259;
      W_o[10,9] := -0.09774768;
      W_o[10,10] := 0.10358307;
      W_o[10,11] := -0.31610432;
      W_o[10,12] := -0.14680047;
      W_o[10,13] := 0.00749488;
      W_o[10,14] := -0.24110141;
      W_o[10,15] := 0.08747873;
      W_o[10,16] := -0.00101395;
      W_o[10,17] := 0.47821096;
      W_o[10,18] := -0.15641819;
      W_o[10,19] := 0.59271890;
      W_o[10,20] := -0.04229831;
      W_o[10,21] := 0.38243753;
      W_o[10,22] := -0.26737732;
      W_o[10,23] := -0.44031852;
      W_o[10,24] := -0.06061750;
      W_o[10,25] := 0.08338970;
      W_o[10,26] := 0.16046619;
      W_o[10,27] := -0.29012343;
      W_o[10,28] := -0.09002028;
      W_o[10,29] := 0.50669360;
      W_o[10,30] := -0.02974824;
      W_o[10,31] := -0.07661217;
      W_o[10,32] := 0.01027904;
      W_o[10,33] := 0.17289472;
      W_o[10,34] := 0.25320745;
      W_o[10,35] := -0.02873696;
      W_o[10,36] := 0.02370308;
      W_o[10,37] := -0.01131884;
      W_o[10,38] := 0.09573818;
      W_o[10,39] := 0.47049189;
      W_o[11,0] := -0.45122087;
      W_o[11,1] := -0.24837552;
      W_o[11,2] := -0.17518084;
      W_o[11,3] := -0.14433257;
      W_o[11,4] := -0.03657356;
      W_o[11,5] := 0.12127155;
      W_o[11,6] := 0.02119773;
      W_o[11,7] := -0.32717624;
      W_o[11,8] := -0.07766484;
      W_o[11,9] := -0.24478522;
      W_o[11,10] := -0.44142914;
      W_o[11,11] := -0.17975523;
      W_o[11,12] := 0.00227619;
      W_o[11,13] := 0.07897434;
      W_o[11,14] := 0.08925162;
      W_o[11,15] := -0.27678323;
      W_o[11,16] := 0.03997169;
      W_o[11,17] := 0.04137829;
      W_o[11,18] := 0.04908814;
      W_o[11,19] := -0.09592513;
      W_o[11,20] := -0.05133458;
      W_o[11,21] := 0.07453518;
      W_o[11,22] := -0.01675062;
      W_o[11,23] := -0.11344488;
      W_o[11,24] := -0.83213097;
      W_o[11,25] := -0.29627800;
      W_o[11,26] := -0.02552608;
      W_o[11,27] := -0.03361585;
      W_o[11,28] := 0.15408768;
      W_o[11,29] := -0.05364017;
      W_o[11,30] := -0.04533393;
      W_o[11,31] := 0.03891878;
      W_o[11,32] := 0.01682842;
      W_o[11,33] := 0.20843782;
      W_o[11,34] := 0.17199376;
      W_o[11,35] := 0.03853744;
      W_o[11,36] := -0.07420836;
      W_o[11,37] := 0.25969163;
      W_o[11,38] := -0.04495483;
      W_o[11,39] := 0.31751272;
      W_o[12,0] := -0.45846713;
      W_o[12,1] := 0.01219229;
      W_o[12,2] := -0.21452378;
      W_o[12,3] := 0.34776640;
      W_o[12,4] := -0.29397878;
      W_o[12,5] := 0.41532251;
      W_o[12,6] := -0.13071139;
      W_o[12,7] := 0.44153231;
      W_o[12,8] := -0.61726791;
      W_o[12,9] := 0.87728906;
      W_o[12,10] := 0.19736496;
      W_o[12,11] := -0.36575502;
      W_o[12,12] := -0.06834572;
      W_o[12,13] := -0.09713604;
      W_o[12,14] := -0.94619924;
      W_o[12,15] := -0.49495792;
      W_o[12,16] := -0.38597691;
      W_o[12,17] := 0.25405318;
      W_o[12,18] := -0.35970402;
      W_o[12,19] := -0.31992292;
      W_o[12,20] := -0.05041254;
      W_o[12,21] := 0.29023391;
      W_o[12,22] := 0.04701138;
      W_o[12,23] := -0.00951147;
      W_o[12,24] := 0.07614060;
      W_o[12,25] := 0.10633016;
      W_o[12,26] := -0.41119781;
      W_o[12,27] := 0.24563172;
      W_o[12,28] := 0.20139630;
      W_o[12,29] := -0.04020792;
      W_o[12,30] := -0.14353402;
      W_o[12,31] := 0.19642521;
      W_o[12,32] := -0.01561482;
      W_o[12,33] := 0.11414265;
      W_o[12,34] := 0.21035014;
      W_o[12,35] := -0.20196043;
      W_o[12,36] := -0.01346343;
      W_o[12,37] := 0.00886301;
      W_o[12,38] := -0.44273621;
      W_o[12,39] := -0.95633447;
      W_o[13,0] := 0.29477751;
      W_o[13,1] := -0.53577411;
      W_o[13,2] := -0.02068770;
      W_o[13,3] := 0.18331867;
      W_o[13,4] := 0.06520753;
      W_o[13,5] := -0.24880944;
      W_o[13,6] := 0.33745202;
      W_o[13,7] := 0.29234564;
      W_o[13,8] := -0.17960128;
      W_o[13,9] := 0.11059473;
      W_o[13,10] := -0.39583328;
      W_o[13,11] := -0.14740023;
      W_o[13,12] := -0.13524790;
      W_o[13,13] := -0.48056528;
      W_o[13,14] := 0.00853791;
      W_o[13,15] := -0.10090394;
      W_o[13,16] := 0.33605260;
      W_o[13,17] := 0.23146117;
      W_o[13,18] := -0.05673217;
      W_o[13,19] := -0.47146145;
      W_o[13,20] := -0.12118670;
      W_o[13,21] := -0.70609426;
      W_o[13,22] := 0.36966327;
      W_o[13,23] := -0.44564933;
      W_o[13,24] := 1.55096805;
      W_o[13,25] := 1.31797290;
      W_o[13,26] := -0.51299953;
      W_o[13,27] := -0.13438945;
      W_o[13,28] := -0.38488221;
      W_o[13,29] := -0.13619691;
      W_o[13,30] := 0.43576846;
      W_o[13,31] := 0.42430091;
      W_o[13,32] := 0.46291351;
      W_o[13,33] := 0.14588232;
      W_o[13,34] := 1.15397358;
      W_o[13,35] := 0.20940591;
      W_o[13,36] := 0.04176854;
      W_o[13,37] := 0.18896750;
      W_o[13,38] := 0.14395012;
      W_o[13,39] := -0.16809192;
      W_o[14,0] := -0.07066596;
      W_o[14,1] := -0.09891939;
      W_o[14,2] := 0.01945558;
      W_o[14,3] := -0.04060903;
      W_o[14,4] := -0.10807311;
      W_o[14,5] := -0.09394543;
      W_o[14,6] := 0.30761227;
      W_o[14,7] := 0.31411666;
      W_o[14,8] := -0.12813382;
      W_o[14,9] := 0.62423646;
      W_o[14,10] := -0.71268511;
      W_o[14,11] := -0.23432153;
      W_o[14,12] := 0.00524576;
      W_o[14,13] := 0.14269492;
      W_o[14,14] := -0.14689596;
      W_o[14,15] := -0.02694557;
      W_o[14,16] := -0.00629303;
      W_o[14,17] := -0.10897459;
      W_o[14,18] := 0.11965847;
      W_o[14,19] := 0.16928390;
      W_o[14,20] := -1.25712538;
      W_o[14,21] := 0.05357262;
      W_o[14,22] := -0.18104394;
      W_o[14,23] := -0.12610403;
      W_o[14,24] := 0.22656150;
      W_o[14,25] := 0.13174540;
      W_o[14,26] := -0.35520098;
      W_o[14,27] := -0.38631681;
      W_o[14,28] := -0.11225829;
      W_o[14,29] := 0.01531188;
      W_o[14,30] := -0.34894708;
      W_o[14,31] := -0.46126148;
      W_o[14,32] := 0.24300313;
      W_o[14,33] := -0.32292667;
      W_o[14,34] := -0.31053829;
      W_o[14,35] := 0.50295210;
      W_o[14,36] := 0.07078700;
      W_o[14,37] := 0.37107170;
      W_o[14,38] := 0.03356927;
      W_o[14,39] := 0.21596275;
      W_o[15,0] := -0.01927980;
      W_o[15,1] := 0.62023401;
      W_o[15,2] := -0.38161528;
      W_o[15,3] := 0.16676347;
      W_o[15,4] := -0.11090784;
      W_o[15,5] := -0.06693771;
      W_o[15,6] := 0.04256647;
      W_o[15,7] := -0.04539243;
      W_o[15,8] := -0.02514778;
      W_o[15,9] := 0.00854907;
      W_o[15,10] := -0.07782564;
      W_o[15,11] := -0.24826944;
      W_o[15,12] := -0.41691181;
      W_o[15,13] := -0.28086716;
      W_o[15,14] := 0.09221611;
      W_o[15,15] := -0.06106566;
      W_o[15,16] := -0.13982905;
      W_o[15,17] := -0.00676943;
      W_o[15,18] := 1.90766096;
      W_o[15,19] := -0.14813134;
      W_o[15,20] := 0.18182682;
      W_o[15,21] := 0.26262483;
      W_o[15,22] := -0.01057434;
      W_o[15,23] := -0.18209115;
      W_o[15,24] := 0.13505831;
      W_o[15,25] := 0.29596528;
      W_o[15,26] := 0.07817908;
      W_o[15,27] := 0.05244986;
      W_o[15,28] := 0.18200800;
      W_o[15,29] := 0.09552819;
      W_o[15,30] := 0.19191824;
      W_o[15,31] := -0.09961358;
      W_o[15,32] := 0.14266075;
      W_o[15,33] := 0.11388518;
      W_o[15,34] := 0.19663931;
      W_o[15,35] := 0.16248274;
      W_o[15,36] := 0.02574501;
      W_o[15,37] := 0.08326160;
      W_o[15,38] := 0.05700103;
      W_o[15,39] := -0.10967547;
      W_o[16,0] := -0.12055943;
      W_o[16,1] := 0.02352543;
      W_o[16,2] := 0.12517351;
      W_o[16,3] := 0.08651733;
      W_o[16,4] := -0.12547506;
      W_o[16,5] := 0.02112064;
      W_o[16,6] := -0.08796533;
      W_o[16,7] := -0.24835224;
      W_o[16,8] := 0.04001724;
      W_o[16,9] := 0.06488604;
      W_o[16,10] := -0.02771191;
      W_o[16,11] := -0.17178981;
      W_o[16,12] := 0.22396629;
      W_o[16,13] := 0.09256334;
      W_o[16,14] := 1.44004285;
      W_o[16,15] := 0.17223491;
      W_o[16,16] := -0.10340090;
      W_o[16,17] := -0.23361848;
      W_o[16,18] := -0.14158271;
      W_o[16,19] := -0.29240519;
      W_o[16,20] := -0.20497365;
      W_o[16,21] := -0.24302354;
      W_o[16,22] := -0.26764143;
      W_o[16,23] := -0.16838124;
      W_o[16,24] := 0.09174137;
      W_o[16,25] := 0.10078798;
      W_o[16,26] := -0.05724070;
      W_o[16,27] := 0.16470623;
      W_o[16,28] := -0.01910415;
      W_o[16,29] := 0.10625532;
      W_o[16,30] := -0.47499156;
      W_o[16,31] := -0.29816622;
      W_o[16,32] := 0.11608597;
      W_o[16,33] := 0.24367557;
      W_o[16,34] := 0.07241584;
      W_o[16,35] := -0.00182753;
      W_o[16,36] := -0.03502716;
      W_o[16,37] := 0.04038282;
      W_o[16,38] := -0.46209079;
      W_o[16,39] := -0.03488237;
      W_o[17,0] := 0.19619699;
      W_o[17,1] := -0.01224999;
      W_o[17,2] := -0.09592830;
      W_o[17,3] := 0.13105205;
      W_o[17,4] := -0.06990813;
      W_o[17,5] := 0.12131099;
      W_o[17,6] := -0.36796319;
      W_o[17,7] := 0.01895757;
      W_o[17,8] := -0.14479473;
      W_o[17,9] := -0.05460491;
      W_o[17,10] := -0.21064177;
      W_o[17,11] := -0.15560260;
      W_o[17,12] := 0.36397913;
      W_o[17,13] := 0.00632168;
      W_o[17,14] := -0.02379812;
      W_o[17,15] := -0.10433174;
      W_o[17,16] := 0.13820401;
      W_o[17,17] := 0.03157768;
      W_o[17,18] := 0.06665690;
      W_o[17,19] := -0.07547057;
      W_o[17,20] := -0.06856900;
      W_o[17,21] := 0.35087839;
      W_o[17,22] := 0.41616750;
      W_o[17,23] := 0.22190954;
      W_o[17,24] := -0.39432350;
      W_o[17,25] := -0.50648206;
      W_o[17,26] := -0.43276054;
      W_o[17,27] := -0.28167576;
      W_o[17,28] := 0.33131412;
      W_o[17,29] := -0.43105629;
      W_o[17,30] := 0.41572836;
      W_o[17,31] := 0.40853822;
      W_o[17,32] := -0.18380405;
      W_o[17,33] := 0.06230948;
      W_o[17,34] := -1.02132106;
      W_o[17,35] := -0.44359389;
      W_o[17,36] := 0.22586185;
      W_o[17,37] := -0.60560203;
      W_o[17,38] := -0.02626733;
      W_o[17,39] := -0.12374443;
      W_o[18,0] := 0.67671382;
      W_o[18,1] := -0.02955803;
      W_o[18,2] := -0.69954222;
      W_o[18,3] := -0.21833202;
      W_o[18,4] := 0.11020873;
      W_o[18,5] := 0.05349873;
      W_o[18,6] := 0.01451667;
      W_o[18,7] := -0.01579341;
      W_o[18,8] := 0.08036178;
      W_o[18,9] := 0.04839315;
      W_o[18,10] := 0.12851113;
      W_o[18,11] := -0.09096859;
      W_o[18,12] := 0.44943687;
      W_o[18,13] := -0.05456711;
      W_o[18,14] := -0.00199916;
      W_o[18,15] := -0.59411538;
      W_o[18,16] := 0.36505663;
      W_o[18,17] := 0.09268996;
      W_o[18,18] := 0.39661846;
      W_o[18,19] := -0.09039351;
      W_o[18,20] := -0.11261550;
      W_o[18,21] := -0.07885239;
      W_o[18,22] := -0.32996053;
      W_o[18,23] := -0.02365809;
      W_o[18,24] := 0.02115683;
      W_o[18,25] := -0.23625188;
      W_o[18,26] := -0.40231401;
      W_o[18,27] := -0.19057028;
      W_o[18,28] := -0.08412448;
      W_o[18,29] := 0.47558784;
      W_o[18,30] := -0.07593910;
      W_o[18,31] := 0.00504192;
      W_o[18,32] := 0.06475038;
      W_o[18,33] := -0.12659657;
      W_o[18,34] := -0.35659128;
      W_o[18,35] := 0.03855544;
      W_o[18,36] := 0.01103517;
      W_o[18,37] := 0.34359896;
      W_o[18,38] := 0.17736463;
      W_o[18,39] := -0.02774378;
      W_o[19,0] := 0.10965693;
      W_o[19,1] := 0.01622399;
      W_o[19,2] := -0.05064026;
      W_o[19,3] := 0.13318102;
      W_o[19,4] := 0.24355040;
      W_o[19,5] := -0.00512605;
      W_o[19,6] := 0.44769040;
      W_o[19,7] := -0.00255203;
      W_o[19,8] := 0.01048099;
      W_o[19,9] := -0.18939705;
      W_o[19,10] := -0.02095573;
      W_o[19,11] := -0.27015504;
      W_o[19,12] := -0.10165944;
      W_o[19,13] := 0.05600982;
      W_o[19,14] := -0.24807528;
      W_o[19,15] := -0.15258515;
      W_o[19,16] := 0.08634272;
      W_o[19,17] := -0.30263221;
      W_o[19,18] := -0.24419874;
      W_o[19,19] := -0.08025812;
      W_o[19,20] := -0.33539948;
      W_o[19,21] := -0.27438563;
      W_o[19,22] := 0.16595660;
      W_o[19,23] := -0.30487317;
      W_o[19,24] := 1.03807557;
      W_o[19,25] := 1.24136472;
      W_o[19,26] := -0.22411491;
      W_o[19,27] := 0.26359200;
      W_o[19,28] := -0.13634011;
      W_o[19,29] := 0.20968179;
      W_o[19,30] := 0.12642498;
      W_o[19,31] := 0.04515914;
      W_o[19,32] := -0.04690970;
      W_o[19,33] := -0.20752276;
      W_o[19,34] := -0.27094910;
      W_o[19,35] := 0.27156648;
      W_o[19,36] := 0.20130572;
      W_o[19,37] := 0.34102762;
      W_o[19,38] := -0.07027919;
      W_o[19,39] := -0.13568473;
      W_o[20,0] := 0.12208430;
      W_o[20,1] := -1.19830549;
      W_o[20,2] := 0.11077505;
      W_o[20,3] := -0.13637088;
      W_o[20,4] := -0.24187416;
      W_o[20,5] := 0.15134950;
      W_o[20,6] := -0.19458446;
      W_o[20,7] := -0.13166124;
      W_o[20,8] := 0.21297050;
      W_o[20,9] := -0.07992186;
      W_o[20,10] := -0.37585995;
      W_o[20,11] := -0.45625314;
      W_o[20,12] := -0.54481548;
      W_o[20,13] := -0.70314580;
      W_o[20,14] := 0.30990425;
      W_o[20,15] := -0.18910754;
      W_o[20,16] := 0.00197922;
      W_o[20,17] := -0.13265780;
      W_o[20,18] := 0.26902235;
      W_o[20,19] := -0.26386663;
      W_o[20,20] := -0.06443398;
      W_o[20,21] := 0.04061922;
      W_o[20,22] := -0.09064165;
      W_o[20,23] := -0.65842748;
      W_o[20,24] := 0.90004557;
      W_o[20,25] := 0.66679513;
      W_o[20,26] := -0.29249567;
      W_o[20,27] := 0.34693053;
      W_o[20,28] := -0.05513572;
      W_o[20,29] := -0.22162925;
      W_o[20,30] := -0.08319939;
      W_o[20,31] := 0.05482560;
      W_o[20,32] := 0.10454668;
      W_o[20,33] := 0.01671114;
      W_o[20,34] := 0.27574286;
      W_o[20,35] := 0.10379709;
      W_o[20,36] := 0.36904472;
      W_o[20,37] := 0.12985463;
      W_o[20,38] := 0.00496099;
      W_o[20,39] := -0.01408813;
      W_o[21,0] := 0.28419283;
      W_o[21,1] := -0.22313316;
      W_o[21,2] := -0.13725317;
      W_o[21,3] := -0.19043419;
      W_o[21,4] := -0.00902355;
      W_o[21,5] := -0.01000001;
      W_o[21,6] := 0.01011608;
      W_o[21,7] := 0.18769735;
      W_o[21,8] := -0.35901442;
      W_o[21,9] := -0.01924971;
      W_o[21,10] := -0.05591933;
      W_o[21,11] := -0.30113551;
      W_o[21,12] := -0.06003612;
      W_o[21,13] := -0.03653869;
      W_o[21,14] := 0.23013163;
      W_o[21,15] := -0.18402654;
      W_o[21,16] := 0.00067009;
      W_o[21,17] := 0.00555752;
      W_o[21,18] := -0.39069557;
      W_o[21,19] := -0.02719967;
      W_o[21,20] := -0.11985504;
      W_o[21,21] := -0.05135375;
      W_o[21,22] := 0.00483708;
      W_o[21,23] := -0.00932395;
      W_o[21,24] := 1.21189833;
      W_o[21,25] := 1.10336173;
      W_o[21,26] := 0.00207484;
      W_o[21,27] := 0.30631572;
      W_o[21,28] := -0.01023949;
      W_o[21,29] := -0.25422829;
      W_o[21,30] := 0.04308288;
      W_o[21,31] := 0.23724382;
      W_o[21,32] := -0.03441579;
      W_o[21,33] := 0.09921884;
      W_o[21,34] := -0.05138595;
      W_o[21,35] := 0.14999114;
      W_o[21,36] := 0.04971470;
      W_o[21,37] := 0.47195190;
      W_o[21,38] := -0.19572517;
      W_o[21,39] := 0.51274788;
      W_o[22,0] := -0.16943602;
      W_o[22,1] := 0.00563010;
      W_o[22,2] := -0.26435009;
      W_o[22,3] := -0.19878975;
      W_o[22,4] := 0.07118692;
      W_o[22,5] := -0.20846748;
      W_o[22,6] := 0.09807133;
      W_o[22,7] := 0.24857411;
      W_o[22,8] := -0.61267197;
      W_o[22,9] := 0.30163637;
      W_o[22,10] := 0.12847048;
      W_o[22,11] := -0.17597947;
      W_o[22,12] := -0.54820406;
      W_o[22,13] := 0.07215662;
      W_o[22,14] := 0.01129225;
      W_o[22,15] := -0.60692477;
      W_o[22,16] := -0.13993593;
      W_o[22,17] := 0.04423706;
      W_o[22,18] := 0.27432024;
      W_o[22,19] := -0.75937098;
      W_o[22,20] := -0.04410430;
      W_o[22,21] := 0.20002785;
      W_o[22,22] := 0.39420721;
      W_o[22,23] := 0.03570565;
      W_o[22,24] := 0.97649997;
      W_o[22,25] := 0.90339136;
      W_o[22,26] := 0.04228690;
      W_o[22,27] := 0.00061381;
      W_o[22,28] := 0.03039532;
      W_o[22,29] := -0.42651707;
      W_o[22,30] := 0.36901113;
      W_o[22,31] := -0.21120797;
      W_o[22,32] := 0.26569346;
      W_o[22,33] := 0.26688823;
      W_o[22,34] := 1.36073279;
      W_o[22,35] := 0.06819707;
      W_o[22,36] := -0.03853309;
      W_o[22,37] := 0.34158346;
      W_o[22,38] := -0.14647880;
      W_o[22,39] := -0.30082840;
      W_o[23,0] := -0.08132017;
      W_o[23,1] := 0.12405463;
      W_o[23,2] := -0.14107077;
      W_o[23,3] := -0.24506845;
      W_o[23,4] := -0.13199361;
      W_o[23,5] := -0.03389445;
      W_o[23,6] := -0.21414556;
      W_o[23,7] := -0.23311256;
      W_o[23,8] := -0.13650194;
      W_o[23,9] := -0.06286883;
      W_o[23,10] := 0.00841143;
      W_o[23,11] := -0.26586533;
      W_o[23,12] := -0.77279711;
      W_o[23,13] := 0.04476917;
      W_o[23,14] := -0.02570722;
      W_o[23,15] := -0.67947555;
      W_o[23,16] := -0.10737889;
      W_o[23,17] := -0.14506733;
      W_o[23,18] := -0.07871757;
      W_o[23,19] := 0.26410311;
      W_o[23,20] := 0.01176897;
      W_o[23,21] := 0.24851997;
      W_o[23,22] := -0.14329612;
      W_o[23,23] := 0.05818005;
      W_o[23,24] := -0.06095537;
      W_o[23,25] := -0.01079577;
      W_o[23,26] := -0.15323734;
      W_o[23,27] := -0.06460467;
      W_o[23,28] := 0.23262998;
      W_o[23,29] := -0.09089681;
      W_o[23,30] := -0.20274188;
      W_o[23,31] := 0.00825220;
      W_o[23,32] := -0.23682141;
      W_o[23,33] := -0.01393911;
      W_o[23,34] := -0.44447368;
      W_o[23,35] := -0.17238432;
      W_o[23,36] := 0.06580907;
      W_o[23,37] := -0.24129888;
      W_o[23,38] := 0.22879821;
      W_o[23,39] := -0.20935446;
      W_o[24,0] := -0.29845297;
      W_o[24,1] := -0.01605594;
      W_o[24,2] := -0.21348783;
      W_o[24,3] := 0.18770167;
      W_o[24,4] := 0.40503550;
      W_o[24,5] := 0.04710687;
      W_o[24,6] := 0.02535505;
      W_o[24,7] := -0.14365837;
      W_o[24,8] := 0.08790880;
      W_o[24,9] := 0.03595916;
      W_o[24,10] := 0.14366116;
      W_o[24,11] := 0.10561820;
      W_o[24,12] := 0.14821514;
      W_o[24,13] := 0.10624322;
      W_o[24,14] := -0.02442249;
      W_o[24,15] := -0.85966212;
      W_o[24,16] := 0.25513664;
      W_o[24,17] := -0.01131127;
      W_o[24,18] := 0.06305917;
      W_o[24,19] := -0.04991962;
      W_o[24,20] := -0.11697821;
      W_o[24,21] := 0.40113649;
      W_o[24,22] := 0.37508291;
      W_o[24,23] := -0.24759673;
      W_o[24,24] := 0.81437260;
      W_o[24,25] := 0.87859291;
      W_o[24,26] := -0.25504032;
      W_o[24,27] := 0.00359953;
      W_o[24,28] := 0.08905714;
      W_o[24,29] := -0.35785756;
      W_o[24,30] := 0.30963099;
      W_o[24,31] := 0.26427326;
      W_o[24,32] := 0.16915745;
      W_o[24,33] := -0.03463329;
      W_o[24,34] := 1.03964126;
      W_o[24,35] := 0.38874447;
      W_o[24,36] := 0.00002758;
      W_o[24,37] := 0.62176007;
      W_o[24,38] := 0.16058211;
      W_o[24,39] := 0.33820599;
      W_o[25,0] := -0.15827869;
      W_o[25,1] := -0.16348077;
      W_o[25,2] := -0.01712869;
      W_o[25,3] := -0.10746691;
      W_o[25,4] := 0.11193889;
      W_o[25,5] := 0.05051835;
      W_o[25,6] := -0.06929888;
      W_o[25,7] := 0.12160345;
      W_o[25,8] := 0.03813792;
      W_o[25,9] := -0.34885547;
      W_o[25,10] := 0.00919252;
      W_o[25,11] := -0.28402808;
      W_o[25,12] := 0.03405061;
      W_o[25,13] := 0.14783855;
      W_o[25,14] := -0.15031821;
      W_o[25,15] := -0.05125191;
      W_o[25,16] := -0.12565699;
      W_o[25,17] := -0.14568239;
      W_o[25,18] := -0.01262960;
      W_o[25,19] := -0.08616017;
      W_o[25,20] := -0.15277006;
      W_o[25,21] := 0.20841888;
      W_o[25,22] := -0.04930439;
      W_o[25,23] := 0.03694082;
      W_o[25,24] := -0.32650331;
      W_o[25,25] := -0.43368715;
      W_o[25,26] := 0.29667246;
      W_o[25,27] := 0.13562424;
      W_o[25,28] := 0.00602539;
      W_o[25,29] := -0.11556970;
      W_o[25,30] := -0.11670647;
      W_o[25,31] := 0.21641117;
      W_o[25,32] := 0.07681312;
      W_o[25,33] := 0.11902311;
      W_o[25,34] := -0.74214745;
      W_o[25,35] := -0.20617647;
      W_o[25,36] := 0.34914330;
      W_o[25,37] := 0.02189142;
      W_o[25,38] := 0.08599351;
      W_o[25,39] := -0.06438139;
      W_o[26,0] := 0.08425111;
      W_o[26,1] := -0.58966690;
      W_o[26,2] := 0.03988224;
      W_o[26,3] := 0.02729935;
      W_o[26,4] := -0.05624046;
      W_o[26,5] := -0.13146318;
      W_o[26,6] := -0.30366996;
      W_o[26,7] := 0.13844973;
      W_o[26,8] := 0.13473816;
      W_o[26,9] := -0.06228542;
      W_o[26,10] := 0.04189111;
      W_o[26,11] := -0.41877472;
      W_o[26,12] := -0.31954202;
      W_o[26,13] := -0.79478008;
      W_o[26,14] := 0.16057940;
      W_o[26,15] := -0.58071166;
      W_o[26,16] := -0.21012735;
      W_o[26,17] := 0.43383101;
      W_o[26,18] := 0.14964466;
      W_o[26,19] := -0.18990019;
      W_o[26,20] := -0.42491710;
      W_o[26,21] := 0.95986062;
      W_o[26,22] := 0.04300608;
      W_o[26,23] := -0.96704936;
      W_o[26,24] := 0.54781920;
      W_o[26,25] := 0.58229166;
      W_o[26,26] := -0.23230726;
      W_o[26,27] := 0.83588123;
      W_o[26,28] := 0.22317052;
      W_o[26,29] := 0.16007505;
      W_o[26,30] := 0.12239722;
      W_o[26,31] := 0.16152382;
      W_o[26,32] := 0.12553506;
      W_o[26,33] := 0.04014284;
      W_o[26,34] := 0.12537505;
      W_o[26,35] := -0.00895806;
      W_o[26,36] := 0.20728289;
      W_o[26,37] := 0.00799836;
      W_o[26,38] := 0.62892807;
      W_o[26,39] := 0.13861158;
      W_o[27,0] := 0.06326006;
      W_o[27,1] := 0.23618595;
      W_o[27,2] := -0.03490672;
      W_o[27,3] := 0.16602454;
      W_o[27,4] := 0.11501915;
      W_o[27,5] := -0.02404143;
      W_o[27,6] := 0.01201760;
      W_o[27,7] := -0.15343736;
      W_o[27,8] := 0.23991169;
      W_o[27,9] := -0.07392941;
      W_o[27,10] := -0.37113866;
      W_o[27,11] := -0.01294172;
      W_o[27,12] := 0.05966742;
      W_o[27,13] := 0.38502872;
      W_o[27,14] := -0.01520643;
      W_o[27,15] := 0.04960250;
      W_o[27,16] := 0.02223091;
      W_o[27,17] := 0.06513891;
      W_o[27,18] := 0.87503552;
      W_o[27,19] := -0.32749546;
      W_o[27,20] := -0.29846638;
      W_o[27,21] := 0.25289643;
      W_o[27,22] := -0.07202611;
      W_o[27,23] := 0.46618357;
      W_o[27,24] := 0.21820667;
      W_o[27,25] := 0.23740523;
      W_o[27,26] := -0.17351545;
      W_o[27,27] := 0.00297986;
      W_o[27,28] := -0.15194261;
      W_o[27,29] := 0.03098265;
      W_o[27,30] := -0.10000996;
      W_o[27,31] := -0.04632366;
      W_o[27,32] := -0.11644848;
      W_o[27,33] := 0.13315183;
      W_o[27,34] := -0.05289400;
      W_o[27,35] := -0.06853411;
      W_o[27,36] := 0.04859332;
      W_o[27,37] := -0.01074729;
      W_o[27,38] := 0.18418956;
      W_o[27,39] := 0.24411875;
      W_o[28,0] := 0.38454545;
      W_o[28,1] := -0.09921691;
      W_o[28,2] := 0.17482130;
      W_o[28,3] := 0.47387001;
      W_o[28,4] := 0.59608668;
      W_o[28,5] := 1.10501480;
      W_o[28,6] := 0.58899385;
      W_o[28,7] := 0.59814161;
      W_o[28,8] := -0.39170471;
      W_o[28,9] := -0.04862360;
      W_o[28,10] := -0.15780824;
      W_o[28,11] := 0.20561603;
      W_o[28,12] := 0.16484201;
      W_o[28,13] := 0.12286928;
      W_o[28,14] := -0.02785882;
      W_o[28,15] := 0.00350319;
      W_o[28,16] := -0.26939300;
      W_o[28,17] := 0.00739435;
      W_o[28,18] := 0.03591748;
      W_o[28,19] := -0.06792951;
      W_o[28,20] := -0.09338012;
      W_o[28,21] := 0.36284494;
      W_o[28,22] := -0.19505034;
      W_o[28,23] := -0.12139830;
      W_o[28,24] := -0.09270825;
      W_o[28,25] := 0.28046516;
      W_o[28,26] := -0.01498493;
      W_o[28,27] := 0.05435069;
      W_o[28,28] := -0.34572619;
      W_o[28,29] := 0.11151223;
      W_o[28,30] := -0.19364205;
      W_o[28,31] := 0.00614947;
      W_o[28,32] := 0.01484237;
      W_o[28,33] := -0.00043672;
      W_o[28,34] := -0.02858257;
      W_o[28,35] := 0.10208395;
      W_o[28,36] := -0.03411613;
      W_o[28,37] := 0.02349477;
      W_o[28,38] := 0.13816315;
      W_o[28,39] := 0.52501553;
      W_o[29,0] := -0.18324779;
      W_o[29,1] := -0.05853816;
      W_o[29,2] := 0.26039451;
      W_o[29,3] := -0.98865104;
      W_o[29,4] := -0.15028648;
      W_o[29,5] := -0.15060133;
      W_o[29,6] := -0.12402279;
      W_o[29,7] := -0.94413263;
      W_o[29,8] := -0.40111613;
      W_o[29,9] := -0.94540298;
      W_o[29,10] := -0.11447112;
      W_o[29,11] := 0.06361326;
      W_o[29,12] := -0.02295774;
      W_o[29,13] := -0.16729216;
      W_o[29,14] := -0.01723751;
      W_o[29,15] := 0.03889744;
      W_o[29,16] := 0.01416754;
      W_o[29,17] := 0.18922821;
      W_o[29,18] := 0.62092680;
      W_o[29,19] := -0.05044166;
      W_o[29,20] := -0.14229977;
      W_o[29,21] := 0.46528375;
      W_o[29,22] := -0.07385064;
      W_o[29,23] := -0.05523294;
      W_o[29,24] := -0.12556942;
      W_o[29,25] := 0.02227050;
      W_o[29,26] := 0.12705496;
      W_o[29,27] := 0.23423049;
      W_o[29,28] := 0.22679651;
      W_o[29,29] := 0.08325709;
      W_o[29,30] := -0.07831824;
      W_o[29,31] := 0.09269150;
      W_o[29,32] := 0.23119086;
      W_o[29,33] := 0.00614441;
      W_o[29,34] := -0.03272606;
      W_o[29,35] := 0.21645607;
      W_o[29,36] := -0.08076635;
      W_o[29,37] := 0.19516927;
      W_o[29,38] := -0.10431720;
      W_o[29,39] := 0.34962577;
      W_o[30,0] := -0.17053279;
      W_o[30,1] := 0.28092715;
      W_o[30,2] := -0.25433207;
      W_o[30,3] := 0.42893410;
      W_o[30,4] := 0.29364955;
      W_o[30,5] := 0.45948777;
      W_o[30,6] := 0.20079698;
      W_o[30,7] := 0.30596188;
      W_o[30,8] := -0.21047817;
      W_o[30,9] := 0.15506689;
      W_o[30,10] := 0.00432611;
      W_o[30,11] := -0.62245870;
      W_o[30,12] := 0.14567345;
      W_o[30,13] := 0.07906670;
      W_o[30,14] := -0.14710122;
      W_o[30,15] := -1.04116786;
      W_o[30,16] := -0.02922401;
      W_o[30,17] := 0.73474240;
      W_o[30,18] := -0.11361318;
      W_o[30,19] := -0.12736081;
      W_o[30,20] := -0.54530185;
      W_o[30,21] := 0.37676060;
      W_o[30,22] := -0.10530942;
      W_o[30,23] := 0.93415534;
      W_o[30,24] := 0.12902859;
      W_o[30,25] := 0.15574846;
      W_o[30,26] := -0.30366293;
      W_o[30,27] := 0.25573662;
      W_o[30,28] := -0.03016189;
      W_o[30,29] := -0.08305828;
      W_o[30,30] := 0.05287048;
      W_o[30,31] := -0.17765103;
      W_o[30,32] := -0.03835172;
      W_o[30,33] := -0.09356602;
      W_o[30,34] := 0.04692689;
      W_o[30,35] := -0.05208236;
      W_o[30,36] := 0.16482487;
      W_o[30,37] := 0.11884566;
      W_o[30,38] := -0.06400402;
      W_o[30,39] := 0.40286413;
      W_o[31,0] := 0.16404290;
      W_o[31,1] := 0.46366262;
      W_o[31,2] := -0.38138533;
      W_o[31,3] := -0.46019378;
      W_o[31,4] := -0.01337012;
      W_o[31,5] := -0.18527511;
      W_o[31,6] := 0.17191447;
      W_o[31,7] := -0.23169285;
      W_o[31,8] := -0.30011240;
      W_o[31,9] := -0.35588530;
      W_o[31,10] := 0.28456184;
      W_o[31,11] := -0.07606647;
      W_o[31,12] := 0.18738757;
      W_o[31,13] := 0.09178647;
      W_o[31,14] := -0.36835101;
      W_o[31,15] := -0.21991540;
      W_o[31,16] := -0.10830630;
      W_o[31,17] := -0.02204164;
      W_o[31,18] := 0.34590438;
      W_o[31,19] := -0.03473870;
      W_o[31,20] := -0.08824793;
      W_o[31,21] := 0.23285167;
      W_o[31,22] := 0.13429588;
      W_o[31,23] := -0.05079326;
      W_o[31,24] := 1.01064575;
      W_o[31,25] := 0.93705499;
      W_o[31,26] := -0.00717605;
      W_o[31,27] := 0.19875413;
      W_o[31,28] := 0.12919939;
      W_o[31,29] := 0.40136379;
      W_o[31,30] := 0.16724311;
      W_o[31,31] := 0.20745699;
      W_o[31,32] := 0.17766902;
      W_o[31,33] := 0.04470662;
      W_o[31,34] := 0.01820830;
      W_o[31,35] := 0.04602371;
      W_o[31,36] := -0.04520386;
      W_o[31,37] := 0.15461211;
      W_o[31,38] := 0.10138816;
      W_o[31,39] := 0.13385615;
      R_i[0,0] := 0.51221442;
      R_i[0,1] := -0.08369232;
      R_i[0,2] := 0.03878905;
      R_i[0,3] := 0.20494133;
      R_i[0,4] := -0.03932563;
      R_i[0,5] := 0.08536161;
      R_i[0,6] := 0.30735824;
      R_i[0,7] := -0.12362177;
      R_i[0,8] := -0.08596776;
      R_i[0,9] := -0.32035100;
      R_i[0,10] := 0.15439482;
      R_i[0,11] := -0.12604460;
      R_i[0,12] := -0.02973188;
      R_i[0,13] := 0.05927557;
      R_i[0,14] := -0.07623336;
      R_i[0,15] := -0.00301596;
      R_i[0,16] := 0.32530278;
      R_i[0,17] := 0.05220976;
      R_i[0,18] := 0.11539400;
      R_i[0,19] := 0.18311976;
      R_i[0,20] := 0.00480020;
      R_i[0,21] := 0.25051382;
      R_i[0,22] := -0.04145733;
      R_i[0,23] := 0.07402290;
      R_i[0,24] := -0.20104395;
      R_i[0,25] := 0.05086588;
      R_i[0,26] := 0.35890043;
      R_i[0,27] := -0.26820049;
      R_i[0,28] := 0.14356384;
      R_i[0,29] := 0.04561891;
      R_i[0,30] := -0.08693960;
      R_i[0,31] := 0.05159991;
      R_i[1,0] := -0.39476180;
      R_i[1,1] := -0.54307437;
      R_i[1,2] := -0.29268599;
      R_i[1,3] := -0.10010588;
      R_i[1,4] := 0.24404499;
      R_i[1,5] := 0.14846084;
      R_i[1,6] := -0.05601619;
      R_i[1,7] := 0.02294470;
      R_i[1,8] := -0.16648757;
      R_i[1,9] := 0.32459068;
      R_i[1,10] := -0.01827455;
      R_i[1,11] := 0.19746210;
      R_i[1,12] := 0.11636473;
      R_i[1,13] := 0.00401034;
      R_i[1,14] := -0.24268822;
      R_i[1,15] := 0.10728395;
      R_i[1,16] := 0.21394157;
      R_i[1,17] := 0.32035813;
      R_i[1,18] := 0.42325589;
      R_i[1,19] := 0.04751065;
      R_i[1,20] := -0.10960548;
      R_i[1,21] := 0.07085693;
      R_i[1,22] := -0.09014911;
      R_i[1,23] := 0.48759651;
      R_i[1,24] := -0.00283297;
      R_i[1,25] := -0.21995039;
      R_i[1,26] := 0.22566356;
      R_i[1,27] := 0.20846392;
      R_i[1,28] := 0.43219981;
      R_i[1,29] := 0.19601935;
      R_i[1,30] := 0.00557092;
      R_i[1,31] := -0.15710679;
      R_i[2,0] := -0.09799560;
      R_i[2,1] := -0.03242979;
      R_i[2,2] := -0.11478028;
      R_i[2,3] := -0.05793334;
      R_i[2,4] := 0.18223813;
      R_i[2,5] := 0.25427604;
      R_i[2,6] := -0.23983784;
      R_i[2,7] := -0.02530777;
      R_i[2,8] := 0.16238339;
      R_i[2,9] := -0.01505891;
      R_i[2,10] := -0.02597539;
      R_i[2,11] := 0.29585776;
      R_i[2,12] := -0.24353874;
      R_i[2,13] := 0.12663041;
      R_i[2,14] := -0.08277308;
      R_i[2,15] := 0.28346336;
      R_i[2,16] := -0.00677738;
      R_i[2,17] := 0.11487118;
      R_i[2,18] := 0.06775200;
      R_i[2,19] := -0.44146669;
      R_i[2,20] := 0.23812422;
      R_i[2,21] := 0.25623590;
      R_i[2,22] := -0.32976091;
      R_i[2,23] := -0.23411497;
      R_i[2,24] := 0.15387745;
      R_i[2,25] := -0.04061436;
      R_i[2,26] := -0.06825281;
      R_i[2,27] := -0.10614515;
      R_i[2,28] := 0.06188334;
      R_i[2,29] := 0.04751145;
      R_i[2,30] := -0.02594229;
      R_i[2,31] := -0.08297227;
      R_i[3,0] := 0.59734422;
      R_i[3,1] := 0.62934798;
      R_i[3,2] := -0.28277254;
      R_i[3,3] := -0.14456962;
      R_i[3,4] := 0.22697103;
      R_i[3,5] := -0.24137557;
      R_i[3,6] := -0.09450015;
      R_i[3,7] := -0.28781146;
      R_i[3,8] := 0.10587214;
      R_i[3,9] := 0.05082055;
      R_i[3,10] := -0.01967472;
      R_i[3,11] := -0.04364250;
      R_i[3,12] := -0.10228609;
      R_i[3,13] := -0.43443522;
      R_i[3,14] := -0.05234408;
      R_i[3,15] := 0.00316776;
      R_i[3,16] := 0.25638989;
      R_i[3,17] := -0.57547498;
      R_i[3,18] := -0.58224237;
      R_i[3,19] := 0.29023883;
      R_i[3,20] := -0.30726695;
      R_i[3,21] := -0.23389202;
      R_i[3,22] := 0.10424740;
      R_i[3,23] := 0.50697947;
      R_i[3,24] := 0.67361164;
      R_i[3,25] := 0.11139195;
      R_i[3,26] := 0.21593073;
      R_i[3,27] := -0.16444562;
      R_i[3,28] := -0.31045249;
      R_i[3,29] := -0.16161352;
      R_i[3,30] := 0.41730696;
      R_i[3,31] := 0.22310457;
      R_i[4,0] := -0.68015325;
      R_i[4,1] := -0.05127423;
      R_i[4,2] := -0.39381805;
      R_i[4,3] := 0.05806528;
      R_i[4,4] := -0.79496628;
      R_i[4,5] := -0.20844424;
      R_i[4,6] := -0.29482576;
      R_i[4,7] := -0.19208500;
      R_i[4,8] := -0.03055103;
      R_i[4,9] := 0.17312987;
      R_i[4,10] := 0.29928619;
      R_i[4,11] := 0.01625600;
      R_i[4,12] := 0.03432601;
      R_i[4,13] := 0.15404135;
      R_i[4,14] := -0.32348749;
      R_i[4,15] := 0.15164973;
      R_i[4,16] := -0.14383729;
      R_i[4,17] := 0.50618845;
      R_i[4,18] := 0.15368445;
      R_i[4,19] := -0.14246292;
      R_i[4,20] := -0.39640063;
      R_i[4,21] := -0.15193579;
      R_i[4,22] := -0.25101894;
      R_i[4,23] := 0.31156206;
      R_i[4,24] := -0.34337518;
      R_i[4,25] := 0.11715125;
      R_i[4,26] := -0.12993719;
      R_i[4,27] := 0.00820147;
      R_i[4,28] := 0.01172253;
      R_i[4,29] := -0.10363425;
      R_i[4,30] := -0.05802570;
      R_i[4,31] := 0.17425007;
      R_i[5,0] := 0.04320075;
      R_i[5,1] := 0.49440038;
      R_i[5,2] := -0.19613867;
      R_i[5,3] := -0.13992621;
      R_i[5,4] := 0.18828946;
      R_i[5,5] := -0.30870205;
      R_i[5,6] := -0.38518646;
      R_i[5,7] := 0.08675630;
      R_i[5,8] := -0.08192702;
      R_i[5,9] := 0.30595222;
      R_i[5,10] := -0.08707682;
      R_i[5,11] := 0.34791610;
      R_i[5,12] := 0.15098788;
      R_i[5,13] := 0.22802135;
      R_i[5,14] := -0.30620182;
      R_i[5,15] := 0.37073833;
      R_i[5,16] := 0.37478310;
      R_i[5,17] := 0.45391643;
      R_i[5,18] := 0.06185832;
      R_i[5,19] := -0.33158338;
      R_i[5,20] := -0.02432890;
      R_i[5,21] := 0.18415853;
      R_i[5,22] := -0.10519998;
      R_i[5,23] := -0.32212982;
      R_i[5,24] := 0.06411852;
      R_i[5,25] := -0.15758936;
      R_i[5,26] := 0.02480984;
      R_i[5,27] := -0.01958706;
      R_i[5,28] := -0.10984096;
      R_i[5,29] := -0.11458004;
      R_i[5,30] := -0.15903004;
      R_i[5,31] := -0.36854565;
      R_i[6,0] := -0.44474992;
      R_i[6,1] := -0.14604338;
      R_i[6,2] := -0.20325679;
      R_i[6,3] := 0.07389074;
      R_i[6,4] := -0.11414720;
      R_i[6,5] := 0.15199620;
      R_i[6,6] := 0.87022948;
      R_i[6,7] := -0.21483621;
      R_i[6,8] := 0.01107073;
      R_i[6,9] := 0.14963895;
      R_i[6,10] := 0.30801591;
      R_i[6,11] := 0.02712611;
      R_i[6,12] := -0.27252647;
      R_i[6,13] := 0.15130866;
      R_i[6,14] := -0.14920071;
      R_i[6,15] := 0.00198815;
      R_i[6,16] := 0.12359401;
      R_i[6,17] := 0.05180132;
      R_i[6,18] := -0.12470315;
      R_i[6,19] := 0.02542710;
      R_i[6,20] := 0.03194568;
      R_i[6,21] := 0.11095844;
      R_i[6,22] := 0.28193268;
      R_i[6,23] := 0.38227135;
      R_i[6,24] := 0.37125403;
      R_i[6,25] := 0.06781208;
      R_i[6,26] := 0.07599112;
      R_i[6,27] := 0.18019117;
      R_i[6,28] := 0.18807802;
      R_i[6,29] := 0.20881404;
      R_i[6,30] := 0.19318885;
      R_i[6,31] := -0.30889073;
      R_i[7,0] := 0.04426930;
      R_i[7,1] := 0.25343812;
      R_i[7,2] := -0.17179920;
      R_i[7,3] := -0.16134921;
      R_i[7,4] := 0.29839942;
      R_i[7,5] := 0.14249474;
      R_i[7,6] := 0.02440364;
      R_i[7,7] := 0.19092458;
      R_i[7,8] := 0.00073451;
      R_i[7,9] := 0.09839897;
      R_i[7,10] := -0.01482648;
      R_i[7,11] := 0.08983578;
      R_i[7,12] := 0.15308072;
      R_i[7,13] := -0.15867147;
      R_i[7,14] := -0.11703056;
      R_i[7,15] := 0.41265205;
      R_i[7,16] := 0.12111750;
      R_i[7,17] := 0.12324470;
      R_i[7,18] := -0.10129975;
      R_i[7,19] := -0.47583267;
      R_i[7,20] := -0.15473907;
      R_i[7,21] := 0.53924632;
      R_i[7,22] := -0.10791501;
      R_i[7,23] := -0.10555386;
      R_i[7,24] := 0.34796754;
      R_i[7,25] := -0.35563490;
      R_i[7,26] := 0.10007861;
      R_i[7,27] := -0.13200946;
      R_i[7,28] := 0.12732220;
      R_i[7,29] := 0.36458585;
      R_i[7,30] := -0.28027585;
      R_i[7,31] := -0.01899707;
      R_i[8,0] := 0.09240616;
      R_i[8,1] := 0.17131865;
      R_i[8,2] := -0.34956303;
      R_i[8,3] := -0.53239042;
      R_i[8,4] := 0.34950057;
      R_i[8,5] := -0.44799775;
      R_i[8,6] := -0.26424530;
      R_i[8,7] := 0.30338514;
      R_i[8,8] := 0.08230431;
      R_i[8,9] := -0.06719685;
      R_i[8,10] := -0.17309690;
      R_i[8,11] := 0.45292673;
      R_i[8,12] := 0.09825447;
      R_i[8,13] := 0.04815003;
      R_i[8,14] := -0.36457637;
      R_i[8,15] := 0.22648472;
      R_i[8,16] := -0.17537273;
      R_i[8,17] := -0.01817195;
      R_i[8,18] := 0.36542943;
      R_i[8,19] := -0.24352296;
      R_i[8,20] := 0.07373296;
      R_i[8,21] := 0.23523478;
      R_i[8,22] := -0.25938845;
      R_i[8,23] := 0.00498532;
      R_i[8,24] := 0.18884458;
      R_i[8,25] := -0.47260910;
      R_i[8,26] := 0.12872651;
      R_i[8,27] := -0.02397963;
      R_i[8,28] := -0.17394602;
      R_i[8,29] := -0.20191373;
      R_i[8,30] := -0.11511500;
      R_i[8,31] := -0.32247952;
      R_i[9,0] := -0.43916357;
      R_i[9,1] := 0.15041128;
      R_i[9,2] := -0.42185432;
      R_i[9,3] := -0.12993184;
      R_i[9,4] := 0.32591265;
      R_i[9,5] := 0.09058974;
      R_i[9,6] := -0.13897957;
      R_i[9,7] := -0.18829496;
      R_i[9,8] := -0.24926165;
      R_i[9,9] := 1.35596073;
      R_i[9,10] := 0.55806267;
      R_i[9,11] := 0.11075085;
      R_i[9,12] := 0.04421957;
      R_i[9,13] := 0.21959196;
      R_i[9,14] := -0.35033441;
      R_i[9,15] := 0.00343219;
      R_i[9,16] := -0.20537409;
      R_i[9,17] := 0.53368264;
      R_i[9,18] := -0.02451989;
      R_i[9,19] := -0.22755532;
      R_i[9,20] := -0.40258268;
      R_i[9,21] := 0.07195293;
      R_i[9,22] := 0.01220069;
      R_i[9,23] := 0.49520347;
      R_i[9,24] := -0.08750314;
      R_i[9,25] := -0.01107999;
      R_i[9,26] := -0.07968686;
      R_i[9,27] := -0.12996809;
      R_i[9,28] := 0.01705114;
      R_i[9,29] := 0.37185794;
      R_i[9,30] := 0.12276196;
      R_i[9,31] := 0.20904543;
      R_i[10,0] := 0.08714745;
      R_i[10,1] := 0.02989326;
      R_i[10,2] := 0.07895342;
      R_i[10,3] := -0.03991391;
      R_i[10,4] := -0.16139822;
      R_i[10,5] := 0.00718968;
      R_i[10,6] := 0.26604277;
      R_i[10,7] := -0.11648100;
      R_i[10,8] := -0.10396011;
      R_i[10,9] := -0.10569390;
      R_i[10,10] := 0.51669079;
      R_i[10,11] := 0.19915892;
      R_i[10,12] := -0.00985841;
      R_i[10,13] := 0.04906809;
      R_i[10,14] := -0.42191544;
      R_i[10,15] := -0.15171689;
      R_i[10,16] := -0.78436285;
      R_i[10,17] := -0.10871010;
      R_i[10,18] := 0.49287951;
      R_i[10,19] := -0.05839600;
      R_i[10,20] := 0.29305947;
      R_i[10,21] := 0.02178851;
      R_i[10,22] := -0.42277884;
      R_i[10,23] := 0.46705118;
      R_i[10,24] := -0.06049981;
      R_i[10,25] := -0.04425887;
      R_i[10,26] := -0.29427859;
      R_i[10,27] := 0.22292905;
      R_i[10,28] := 0.23763067;
      R_i[10,29] := 0.10558424;
      R_i[10,30] := -0.27244172;
      R_i[10,31] := -0.14848375;
      R_i[11,0] := -0.20009324;
      R_i[11,1] := 0.22914931;
      R_i[11,2] := -0.08989751;
      R_i[11,3] := -0.52993345;
      R_i[11,4] := 0.20788677;
      R_i[11,5] := -0.32998398;
      R_i[11,6] := -0.11127269;
      R_i[11,7] := -0.17718190;
      R_i[11,8] := -0.18657120;
      R_i[11,9] := 0.28600550;
      R_i[11,10] := 0.09621530;
      R_i[11,11] := 0.74793410;
      R_i[11,12] := 0.00333306;
      R_i[11,13] := -0.01473215;
      R_i[11,14] := -0.53499997;
      R_i[11,15] := 0.07715688;
      R_i[11,16] := -0.25301683;
      R_i[11,17] := 0.33122754;
      R_i[11,18] := -0.15208751;
      R_i[11,19] := -0.14227772;
      R_i[11,20] := -0.13599677;
      R_i[11,21] := 0.01813499;
      R_i[11,22] := -0.11655468;
      R_i[11,23] := 0.09607781;
      R_i[11,24] := 0.14136216;
      R_i[11,25] := 0.17874435;
      R_i[11,26] := 0.20932396;
      R_i[11,27] := -0.09231541;
      R_i[11,28] := 0.16655394;
      R_i[11,29] := -0.07641463;
      R_i[11,30] := -0.35409757;
      R_i[11,31] := 0.09594071;
      R_i[12,0] := -0.11654998;
      R_i[12,1] := 0.26751649;
      R_i[12,2] := 0.22307423;
      R_i[12,3] := -0.07999243;
      R_i[12,4] := -0.02321325;
      R_i[12,5] := 0.05414648;
      R_i[12,6] := -0.15591401;
      R_i[12,7] := -0.26203060;
      R_i[12,8] := -0.58493954;
      R_i[12,9] := -0.02167135;
      R_i[12,10] := 0.12806118;
      R_i[12,11] := -0.02724883;
      R_i[12,12] := -0.58108002;
      R_i[12,13] := -0.19241558;
      R_i[12,14] := -0.09912304;
      R_i[12,15] := 0.17238013;
      R_i[12,16] := 0.09443929;
      R_i[12,17] := 0.16614071;
      R_i[12,18] := -0.18041192;
      R_i[12,19] := 0.08594200;
      R_i[12,20] := 0.18258996;
      R_i[12,21] := 0.09522452;
      R_i[12,22] := 0.41028434;
      R_i[12,23] := -0.28717035;
      R_i[12,24] := 0.02750145;
      R_i[12,25] := 0.32911661;
      R_i[12,26] := 0.04212489;
      R_i[12,27] := 0.40236855;
      R_i[12,28] := -0.10092562;
      R_i[12,29] := 0.64539850;
      R_i[12,30] := 0.52788371;
      R_i[12,31] := -0.75803000;
      R_i[13,0] := -0.39125809;
      R_i[13,1] := 0.05575472;
      R_i[13,2] := -0.03408769;
      R_i[13,3] := -0.15652266;
      R_i[13,4] := -0.16123737;
      R_i[13,5] := 0.24292000;
      R_i[13,6] := -0.30130127;
      R_i[13,7] := -0.24130024;
      R_i[13,8] := 0.00776500;
      R_i[13,9] := 0.11403982;
      R_i[13,10] := 0.09043195;
      R_i[13,11] := -0.07317566;
      R_i[13,12] := -0.40591890;
      R_i[13,13] := 0.32489985;
      R_i[13,14] := -0.20800115;
      R_i[13,15] := 0.00221067;
      R_i[13,16] := -0.10147334;
      R_i[13,17] := -0.24813145;
      R_i[13,18] := 0.03474638;
      R_i[13,19] := -0.18104817;
      R_i[13,20] := 0.28191370;
      R_i[13,21] := 0.10907030;
      R_i[13,22] := -0.33868816;
      R_i[13,23] := -0.01885714;
      R_i[13,24] := 0.29839468;
      R_i[13,25] := 0.10087272;
      R_i[13,26] := -0.01320497;
      R_i[13,27] := 0.06962156;
      R_i[13,28] := -0.11318398;
      R_i[13,29] := 0.18922725;
      R_i[13,30] := 0.09005125;
      R_i[13,31] := -0.30306169;
      R_i[14,0] := 0.01120466;
      R_i[14,1] := 0.11350589;
      R_i[14,2] := -0.23733518;
      R_i[14,3] := 0.35504350;
      R_i[14,4] := 0.42941424;
      R_i[14,5] := -0.35159039;
      R_i[14,6] := 0.01117469;
      R_i[14,7] := -0.11143109;
      R_i[14,8] := 0.44690257;
      R_i[14,9] := 0.12703660;
      R_i[14,10] := -0.11827330;
      R_i[14,11] := 0.02845767;
      R_i[14,12] := -0.25289932;
      R_i[14,13] := 0.18736526;
      R_i[14,14] := 0.77491051;
      R_i[14,15] := 0.23110941;
      R_i[14,16] := 0.21939375;
      R_i[14,17] := -0.24036950;
      R_i[14,18] := -0.17610160;
      R_i[14,19] := -0.37820250;
      R_i[14,20] := 0.52524704;
      R_i[14,21] := -0.12975010;
      R_i[14,22] := 0.16990341;
      R_i[14,23] := -0.30200759;
      R_i[14,24] := -0.05411242;
      R_i[14,25] := 0.35907966;
      R_i[14,26] := -0.27149668;
      R_i[14,27] := -0.05471592;
      R_i[14,28] := -0.05388270;
      R_i[14,29] := -0.40745988;
      R_i[14,30] := 0.23365912;
      R_i[14,31] := 0.33957499;
      R_i[15,0] := 0.16775908;
      R_i[15,1] := 0.07096732;
      R_i[15,2] := -0.04280357;
      R_i[15,3] := 0.30321899;
      R_i[15,4] := -0.11642423;
      R_i[15,5] := 0.18614328;
      R_i[15,6] := 0.48792782;
      R_i[15,7] := 0.09495277;
      R_i[15,8] := -0.01985801;
      R_i[15,9] := 0.14887144;
      R_i[15,10] := 0.15832083;
      R_i[15,11] := -0.16339642;
      R_i[15,12] := 0.28504267;
      R_i[15,13] := -0.04822541;
      R_i[15,14] := -0.06426991;
      R_i[15,15] := -0.64180833;
      R_i[15,16] := 0.13660328;
      R_i[15,17] := 0.24940038;
      R_i[15,18] := 0.13910303;
      R_i[15,19] := -0.02350211;
      R_i[15,20] := -0.04269773;
      R_i[15,21] := -0.02816851;
      R_i[15,22] := 0.15895598;
      R_i[15,23] := 0.16843884;
      R_i[15,24] := 0.16463809;
      R_i[15,25] := -0.01168484;
      R_i[15,26] := -0.02309109;
      R_i[15,27] := -0.20655718;
      R_i[15,28] := 0.09094330;
      R_i[15,29] := -0.04085297;
      R_i[15,30] := -0.08570669;
      R_i[15,31] := -0.05749578;
      R_i[16,0] := 0.13447514;
      R_i[16,1] := -0.01801078;
      R_i[16,2] := -0.05059633;
      R_i[16,3] := -0.08663934;
      R_i[16,4] := 0.00052052;
      R_i[16,5] := 0.34696624;
      R_i[16,6] := 0.44769460;
      R_i[16,7] := 0.03157200;
      R_i[16,8] := -0.44279256;
      R_i[16,9] := -0.14010711;
      R_i[16,10] := 0.65262598;
      R_i[16,11] := 0.22846895;
      R_i[16,12] := -0.53771132;
      R_i[16,13] := 0.00055600;
      R_i[16,14] := 0.17123872;
      R_i[16,15] := 0.17721201;
      R_i[16,16] := 1.09687459;
      R_i[16,17] := -0.17730564;
      R_i[16,18] := -0.08602641;
      R_i[16,19] := -0.08945292;
      R_i[16,20] := 0.12588546;
      R_i[16,21] := -0.43724018;
      R_i[16,22] := -0.58790159;
      R_i[16,23] := 0.30984837;
      R_i[16,24] := -0.30069503;
      R_i[16,25] := 0.27324480;
      R_i[16,26] := 0.03958173;
      R_i[16,27] := -0.27124757;
      R_i[16,28] := 0.42478165;
      R_i[16,29] := 0.03367740;
      R_i[16,30] := -0.14776608;
      R_i[16,31] := -0.16438708;
      R_i[17,0] := 0.05412322;
      R_i[17,1] := 0.33582243;
      R_i[17,2] := -0.28220329;
      R_i[17,3] := -0.49404711;
      R_i[17,4] := 0.76758504;
      R_i[17,5] := -0.49188408;
      R_i[17,6] := 0.35752013;
      R_i[17,7] := -0.02469994;
      R_i[17,8] := 0.01132120;
      R_i[17,9] := 0.66087836;
      R_i[17,10] := 0.68969095;
      R_i[17,11] := -0.20370367;
      R_i[17,12] := 0.48326203;
      R_i[17,13] := -0.96083552;
      R_i[17,14] := -0.78994125;
      R_i[17,15] := 0.91829079;
      R_i[17,16] := -0.23014545;
      R_i[17,17] := -0.56922269;
      R_i[17,18] := 0.03208271;
      R_i[17,19] := -0.26753226;
      R_i[17,20] := 0.46724734;
      R_i[17,21] := -0.25534356;
      R_i[17,22] := 0.55033535;
      R_i[17,23] := 0.10821555;
      R_i[17,24] := 0.27335948;
      R_i[17,25] := -0.07342362;
      R_i[17,26] := 0.13944507;
      R_i[17,27] := -0.22517696;
      R_i[17,28] := -0.94890118;
      R_i[17,29] := -0.01491523;
      R_i[17,30] := 0.22817695;
      R_i[17,31] := 0.14350086;
      R_i[18,0] := -0.08198392;
      R_i[18,1] := 0.08573992;
      R_i[18,2] := 0.12008911;
      R_i[18,3] := -0.13298780;
      R_i[18,4] := -0.16758575;
      R_i[18,5] := 0.24653280;
      R_i[18,6] := 0.01826797;
      R_i[18,7] := 0.27076790;
      R_i[18,8] := -0.35665849;
      R_i[18,9] := 0.02654203;
      R_i[18,10] := -0.17872359;
      R_i[18,11] := -0.03283141;
      R_i[18,12] := -0.43551093;
      R_i[18,13] := -0.17177245;
      R_i[18,14] := -0.13806683;
      R_i[18,15] := 0.09106231;
      R_i[18,16] := -0.08847328;
      R_i[18,17] := 0.35300431;
      R_i[18,18] := 1.28586066;
      R_i[18,19] := -0.16597459;
      R_i[18,20] := 0.07983273;
      R_i[18,21] := 0.02233933;
      R_i[18,22] := 0.06625325;
      R_i[18,23] := 0.27211902;
      R_i[18,24] := -0.17268898;
      R_i[18,25] := 0.22699259;
      R_i[18,26] := -0.25373802;
      R_i[18,27] := -0.13492379;
      R_i[18,28] := 0.03534929;
      R_i[18,29] := 0.26698029;
      R_i[18,30] := 0.21760662;
      R_i[18,31] := -0.02662387;
      R_i[19,0] := 0.15502211;
      R_i[19,1] := 0.03973338;
      R_i[19,2] := -0.32049409;
      R_i[19,3] := -0.05688509;
      R_i[19,4] := -0.17240311;
      R_i[19,5] := -0.16044626;
      R_i[19,6] := 0.00450565;
      R_i[19,7] := 0.28525978;
      R_i[19,8] := -0.08821966;
      R_i[19,9] := 0.11336405;
      R_i[19,10] := 0.07316364;
      R_i[19,11] := -0.05398195;
      R_i[19,12] := 0.21548112;
      R_i[19,13] := -0.04186272;
      R_i[19,14] := -0.28405803;
      R_i[19,15] := 0.02832769;
      R_i[19,16] := 0.23835751;
      R_i[19,17] := 0.25204211;
      R_i[19,18] := 0.10707825;
      R_i[19,19] := -0.31347281;
      R_i[19,20] := 0.26063022;
      R_i[19,21] := 0.42351454;
      R_i[19,22] := -0.13583225;
      R_i[19,23] := 0.22939259;
      R_i[19,24] := -0.21873315;
      R_i[19,25] := -0.22747228;
      R_i[19,26] := -0.10111309;
      R_i[19,27] := -0.33270133;
      R_i[19,28] := -0.20719844;
      R_i[19,29] := 0.15941210;
      R_i[19,30] := 0.05134924;
      R_i[19,31] := -0.05631643;
      R_i[20,0] := -0.00901746;
      R_i[20,1] := 0.06032126;
      R_i[20,2] := -0.22463125;
      R_i[20,3] := -0.07069563;
      R_i[20,4] := -0.47293216;
      R_i[20,5] := 0.06162272;
      R_i[20,6] := 0.04380284;
      R_i[20,7] := -0.20195602;
      R_i[20,8] := 0.52933151;
      R_i[20,9] := 0.17288506;
      R_i[20,10] := 0.09337651;
      R_i[20,11] := -0.26854435;
      R_i[20,12] := 0.04588911;
      R_i[20,13] := -0.09455147;
      R_i[20,14] := -0.17151232;
      R_i[20,15] := -0.33518133;
      R_i[20,16] := 0.14887759;
      R_i[20,17] := 0.10844737;
      R_i[20,18] := 0.03363106;
      R_i[20,19] := -0.18901934;
      R_i[20,20] := -0.37031725;
      R_i[20,21] := 0.17756981;
      R_i[20,22] := -0.09798433;
      R_i[20,23] := -0.25045586;
      R_i[20,24] := 0.26002321;
      R_i[20,25] := -0.25486484;
      R_i[20,26] := -0.00880880;
      R_i[20,27] := 0.27573004;
      R_i[20,28] := 0.05462186;
      R_i[20,29] := -0.06694781;
      R_i[20,30] := -0.37804615;
      R_i[20,31] := -0.56364352;
      R_i[21,0] := 0.03798443;
      R_i[21,1] := -0.11627547;
      R_i[21,2] := -0.38938740;
      R_i[21,3] := -0.03386816;
      R_i[21,4] := 0.34411737;
      R_i[21,5] := -0.31639281;
      R_i[21,6] := -0.17763256;
      R_i[21,7] := -0.02297345;
      R_i[21,8] := 0.07765912;
      R_i[21,9] := 0.15951294;
      R_i[21,10] := 0.65718466;
      R_i[21,11] := -0.17887022;
      R_i[21,12] := -0.03618487;
      R_i[21,13] := -0.06913149;
      R_i[21,14] := 0.18947972;
      R_i[21,15] := 0.07929875;
      R_i[21,16] := -0.04257125;
      R_i[21,17] := -0.18183275;
      R_i[21,18] := -0.13432932;
      R_i[21,19] := 0.24196239;
      R_i[21,20] := -0.14389262;
      R_i[21,21] := 0.88659251;
      R_i[21,22] := 0.23105976;
      R_i[21,23] := -0.00900477;
      R_i[21,24] := 0.29885840;
      R_i[21,25] := 0.54741335;
      R_i[21,26] := 0.20832890;
      R_i[21,27] := -0.67173117;
      R_i[21,28] := 0.06925270;
      R_i[21,29] := -0.02693848;
      R_i[21,30] := -0.20997405;
      R_i[21,31] := 0.23705347;
      R_i[22,0] := -0.12260506;
      R_i[22,1] := 0.10777262;
      R_i[22,2] := -0.29853928;
      R_i[22,3] := -0.15479548;
      R_i[22,4] := 0.30029958;
      R_i[22,5] := -0.02772681;
      R_i[22,6] := 0.31630555;
      R_i[22,7] := -0.21110223;
      R_i[22,8] := 0.39206710;
      R_i[22,9] := -0.27248287;
      R_i[22,10] := -0.32923529;
      R_i[22,11] := 0.35362753;
      R_i[22,12] := -0.13532224;
      R_i[22,13] := -0.35496590;
      R_i[22,14] := -0.00508518;
      R_i[22,15] := 0.05788676;
      R_i[22,16] := 0.03263550;
      R_i[22,17] := 0.12816045;
      R_i[22,18] := 0.19306229;
      R_i[22,19] := -0.26334158;
      R_i[22,20] := -0.33350593;
      R_i[22,21] := -0.02586301;
      R_i[22,22] := 0.36985421;
      R_i[22,23] := -0.05025383;
      R_i[22,24] := 0.13873249;
      R_i[22,25] := 0.05488453;
      R_i[22,26] := 0.10486135;
      R_i[22,27] := -0.08153543;
      R_i[22,28] := 0.50797367;
      R_i[22,29] := 0.13860652;
      R_i[22,30] := -0.01046087;
      R_i[22,31] := -0.40905952;
      R_i[23,0] := 0.03703520;
      R_i[23,1] := 0.35561198;
      R_i[23,2] := -0.15956397;
      R_i[23,3] := 0.06172862;
      R_i[23,4] := -0.00924198;
      R_i[23,5] := -0.30205476;
      R_i[23,6] := 0.35665691;
      R_i[23,7] := 0.02458556;
      R_i[23,8] := -0.07570854;
      R_i[23,9] := 0.21206109;
      R_i[23,10] := 0.06857381;
      R_i[23,11] := 0.29381767;
      R_i[23,12] := -0.05752667;
      R_i[23,13] := 0.01229799;
      R_i[23,14] := 0.02933831;
      R_i[23,15] := 0.17395060;
      R_i[23,16] := 0.19358973;
      R_i[23,17] := 0.30012521;
      R_i[23,18] := -0.20486185;
      R_i[23,19] := -0.07677986;
      R_i[23,20] := -0.10174387;
      R_i[23,21] := 0.02195450;
      R_i[23,22] := -0.03289494;
      R_i[23,23] := 1.05171776;
      R_i[23,24] := 0.34484801;
      R_i[23,25] := 0.14438485;
      R_i[23,26] := 0.17363730;
      R_i[23,27] := 0.04493184;
      R_i[23,28] := 0.37233853;
      R_i[23,29] := 0.07609949;
      R_i[23,30] := 0.30364865;
      R_i[23,31] := -0.14013796;
      R_i[24,0] := 0.34240055;
      R_i[24,1] := -0.14468294;
      R_i[24,2] := -0.31550655;
      R_i[24,3] := -0.13977182;
      R_i[24,4] := -0.20417063;
      R_i[24,5] := 0.16776828;
      R_i[24,6] := 0.02561445;
      R_i[24,7] := -0.05868829;
      R_i[24,8] := -0.02827646;
      R_i[24,9] := 0.19114552;
      R_i[24,10] := -0.15757357;
      R_i[24,11] := 0.26007780;
      R_i[24,12] := 0.21217065;
      R_i[24,13] := 0.13858628;
      R_i[24,14] := 0.00071470;
      R_i[24,15] := -0.15069637;
      R_i[24,16] := 0.29770842;
      R_i[24,17] := 0.16526395;
      R_i[24,18] := -0.15285577;
      R_i[24,19] := -0.18742292;
      R_i[24,20] := -0.06594079;
      R_i[24,21] := -0.04290878;
      R_i[24,22] := -0.25888646;
      R_i[24,23] := -0.12326243;
      R_i[24,24] := 0.25272989;
      R_i[24,25] := -0.20074646;
      R_i[24,26] := 0.12650153;
      R_i[24,27] := -0.30788255;
      R_i[24,28] := 0.20032974;
      R_i[24,29] := 0.13566294;
      R_i[24,30] := -0.09083051;
      R_i[24,31] := -0.14403652;
      R_i[25,0] := -0.00364695;
      R_i[25,1] := 0.06404819;
      R_i[25,2] := -0.01804773;
      R_i[25,3] := 0.04540015;
      R_i[25,4] := 0.16974008;
      R_i[25,5] := -0.08127178;
      R_i[25,6] := 0.19735654;
      R_i[25,7] := -0.08230321;
      R_i[25,8] := -0.37761867;
      R_i[25,9] := 0.12201649;
      R_i[25,10] := 0.10528291;
      R_i[25,11] := -0.10855001;
      R_i[25,12] := 0.23163250;
      R_i[25,13] := -0.12369552;
      R_i[25,14] := -0.21644136;
      R_i[25,15] := 0.28066093;
      R_i[25,16] := -0.00126031;
      R_i[25,17] := 0.34386733;
      R_i[25,18] := -0.05251693;
      R_i[25,19] := 0.11943450;
      R_i[25,20] := 0.12946576;
      R_i[25,21] := 0.32350007;
      R_i[25,22] := -0.16389352;
      R_i[25,23] := 0.06864835;
      R_i[25,24] := -0.02653339;
      R_i[25,25] := 0.44217756;
      R_i[25,26] := -0.21659601;
      R_i[25,27] := -0.06462156;
      R_i[25,28] := 0.14042386;
      R_i[25,29] := 0.25927311;
      R_i[25,30] := -0.08044507;
      R_i[25,31] := -0.20894651;
      R_i[26,0] := -0.25971705;
      R_i[26,1] := 0.07879175;
      R_i[26,2] := 0.11486167;
      R_i[26,3] := 0.03312163;
      R_i[26,4] := -0.31499544;
      R_i[26,5] := 0.22103539;
      R_i[26,6] := 0.60527152;
      R_i[26,7] := 0.12882712;
      R_i[26,8] := 0.03168129;
      R_i[26,9] := 0.34555426;
      R_i[26,10] := 0.20023961;
      R_i[26,11] := 0.00272711;
      R_i[26,12] := 0.59746903;
      R_i[26,13] := 0.15487805;
      R_i[26,14] := 0.00623762;
      R_i[26,15] := 0.10250810;
      R_i[26,16] := 0.29433212;
      R_i[26,17] := 0.48321578;
      R_i[26,18] := 0.34317333;
      R_i[26,19] := 0.10681155;
      R_i[26,20] := -0.23560931;
      R_i[26,21] := 0.16572604;
      R_i[26,22] := -0.30539343;
      R_i[26,23] := 0.02724703;
      R_i[26,24] := -0.11780143;
      R_i[26,25] := -0.25815722;
      R_i[26,26] := 0.34590581;
      R_i[26,27] := -0.34810752;
      R_i[26,28] := 0.06762858;
      R_i[26,29] := -0.09515713;
      R_i[26,30] := 0.14459436;
      R_i[26,31] := -0.25349867;
      R_i[27,0] := 0.03371919;
      R_i[27,1] := -0.04406705;
      R_i[27,2] := -0.24740066;
      R_i[27,3] := -0.61750942;
      R_i[27,4] := -0.03851713;
      R_i[27,5] := 0.20272811;
      R_i[27,6] := 0.04261627;
      R_i[27,7] := -0.63512993;
      R_i[27,8] := 0.07641039;
      R_i[27,9] := 0.08821981;
      R_i[27,10] := -0.07666441;
      R_i[27,11] := 0.20226212;
      R_i[27,12] := -0.58091104;
      R_i[27,13] := -0.29244682;
      R_i[27,14] := -0.32245147;
      R_i[27,15] := 0.58181006;
      R_i[27,16] := -0.39972940;
      R_i[27,17] := 0.21634744;
      R_i[27,18] := 0.48655644;
      R_i[27,19] := 0.10145795;
      R_i[27,20] := 0.06825342;
      R_i[27,21] := 0.01775364;
      R_i[27,22] := 0.48730814;
      R_i[27,23] := 0.03193397;
      R_i[27,24] := 0.20350280;
      R_i[27,25] := -0.08388541;
      R_i[27,26] := -0.37410170;
      R_i[27,27] := 1.49699283;
      R_i[27,28] := 0.00160924;
      R_i[27,29] := 0.25602624;
      R_i[27,30] := 0.35360309;
      R_i[27,31] := -0.48147491;
      R_i[28,0] := 0.16041149;
      R_i[28,1] := -0.11364735;
      R_i[28,2] := 0.20443638;
      R_i[28,3] := -0.25905165;
      R_i[28,4] := 0.32468283;
      R_i[28,5] := -0.16589360;
      R_i[28,6] := 0.02469636;
      R_i[28,7] := -0.44379267;
      R_i[28,8] := -0.16905288;
      R_i[28,9] := 0.34305990;
      R_i[28,10] := -0.17373589;
      R_i[28,11] := 0.01532834;
      R_i[28,12] := 0.17097749;
      R_i[28,13] := -0.36091733;
      R_i[28,14] := -0.12726678;
      R_i[28,15] := -0.13177131;
      R_i[28,16] := -0.03381614;
      R_i[28,17] := 0.57329458;
      R_i[28,18] := 0.10554976;
      R_i[28,19] := -0.48848552;
      R_i[28,20] := 0.01206277;
      R_i[28,21] := -0.01500845;
      R_i[28,22] := -0.10783848;
      R_i[28,23] := -0.14017676;
      R_i[28,24] := 0.11403215;
      R_i[28,25] := -0.02840269;
      R_i[28,26] := 0.41083917;
      R_i[28,27] := 0.03614673;
      R_i[28,28] := 0.90944064;
      R_i[28,29] := 0.17652564;
      R_i[28,30] := -0.66777414;
      R_i[28,31] := -0.43163636;
      R_i[29,0] := -0.05349075;
      R_i[29,1] := -0.12321150;
      R_i[29,2] := 0.06346910;
      R_i[29,3] := -0.38304222;
      R_i[29,4] := 0.34138668;
      R_i[29,5] := 0.08186229;
      R_i[29,6] := 0.12306959;
      R_i[29,7] := -0.18967490;
      R_i[29,8] := 0.15568839;
      R_i[29,9] := 0.16008142;
      R_i[29,10] := 0.07354110;
      R_i[29,11] := 0.23890246;
      R_i[29,12] := 0.32625028;
      R_i[29,13] := 0.27283725;
      R_i[29,14] := -0.38482612;
      R_i[29,15] := -0.08214376;
      R_i[29,16] := 0.03451258;
      R_i[29,17] := 0.53154832;
      R_i[29,18] := 0.32419375;
      R_i[29,19] := 0.08637193;
      R_i[29,20] := -0.23812342;
      R_i[29,21] := -0.12626043;
      R_i[29,22] := -0.20393825;
      R_i[29,23] := 0.41695753;
      R_i[29,24] := -0.03135362;
      R_i[29,25] := -0.09947015;
      R_i[29,26] := 0.19810902;
      R_i[29,27] := -0.07402156;
      R_i[29,28] := -0.23810703;
      R_i[29,29] := 0.26977152;
      R_i[29,30] := -0.22404684;
      R_i[29,31] := 0.17006949;
      R_i[30,0] := 0.03638737;
      R_i[30,1] := 0.05191260;
      R_i[30,2] := -0.52651483;
      R_i[30,3] := -0.86915576;
      R_i[30,4] := -0.15424719;
      R_i[30,5] := -0.21525031;
      R_i[30,6] := 1.08992696;
      R_i[30,7] := -0.20518234;
      R_i[30,8] := 1.81346786;
      R_i[30,9] := -0.30627471;
      R_i[30,10] := 0.27207708;
      R_i[30,11] := 0.15125890;
      R_i[30,12] := -0.37401557;
      R_i[30,13] := -0.13959804;
      R_i[30,14] := -0.01365140;
      R_i[30,15] := 0.04396977;
      R_i[30,16] := 0.32709506;
      R_i[30,17] := -0.88627982;
      R_i[30,18] := -0.37619492;
      R_i[30,19] := -0.09723003;
      R_i[30,20] := -0.29918641;
      R_i[30,21] := -0.43405920;
      R_i[30,22] := -0.10127983;
      R_i[30,23] := 0.23152281;
      R_i[30,24] := 1.14722586;
      R_i[30,25] := -0.13771860;
      R_i[30,26] := -0.59857517;
      R_i[30,27] := -0.38145676;
      R_i[30,28] := -0.11991661;
      R_i[30,29] := 0.40799883;
      R_i[30,30] := -1.59745562;
      R_i[30,31] := -0.37564871;
      R_i[31,0] := -0.05862521;
      R_i[31,1] := -0.03135950;
      R_i[31,2] := -0.55573916;
      R_i[31,3] := -0.13187377;
      R_i[31,4] := 0.34288785;
      R_i[31,5] := 0.30176958;
      R_i[31,6] := 0.31988955;
      R_i[31,7] := -0.13703822;
      R_i[31,8] := 0.25901517;
      R_i[31,9] := 0.41554999;
      R_i[31,10] := -0.34672722;
      R_i[31,11] := -0.21812697;
      R_i[31,12] := -0.13724922;
      R_i[31,13] := -0.27975926;
      R_i[31,14] := -0.46450689;
      R_i[31,15] := 0.07930830;
      R_i[31,16] := -0.04665133;
      R_i[31,17] := 0.59159482;
      R_i[31,18] := -0.07420903;
      R_i[31,19] := -0.13947521;
      R_i[31,20] := 0.02244737;
      R_i[31,21] := 0.18911299;
      R_i[31,22] := 0.41634119;
      R_i[31,23] := 0.14076699;
      R_i[31,24] := 0.40610394;
      R_i[31,25] := -0.39880338;
      R_i[31,26] := -0.25052059;
      R_i[31,27] := -0.13714445;
      R_i[31,28] := 0.26395574;
      R_i[31,29] := -0.31718644;
      R_i[31,30] := -0.14742820;
      R_i[31,31] := -0.38917819;
      R_f[0,0] := 0.67188150;
      R_f[0,1] := 0.34223723;
      R_f[0,2] := 0.18857408;
      R_f[0,3] := -0.07556254;
      R_f[0,4] := 0.21652593;
      R_f[0,5] := -0.06935426;
      R_f[0,6] := -0.09358843;
      R_f[0,7] := 0.04287541;
      R_f[0,8] := 0.13322420;
      R_f[0,9] := 0.06833595;
      R_f[0,10] := -0.42965809;
      R_f[0,11] := -0.05324866;
      R_f[0,12] := -0.07535404;
      R_f[0,13] := -0.05255458;
      R_f[0,14] := 0.49930987;
      R_f[0,15] := -0.18491820;
      R_f[0,16] := 0.11946521;
      R_f[0,17] := -0.75537163;
      R_f[0,18] := -0.02437763;
      R_f[0,19] := 0.13815457;
      R_f[0,20] := -0.16969654;
      R_f[0,21] := 0.03172547;
      R_f[0,22] := 0.17337099;
      R_f[0,23] := -0.25701371;
      R_f[0,24] := -0.12645802;
      R_f[0,25] := 0.10932370;
      R_f[0,26] := 0.02822654;
      R_f[0,27] := -0.00966967;
      R_f[0,28] := -0.09048105;
      R_f[0,29] := 0.00988982;
      R_f[0,30] := 0.10447063;
      R_f[0,31] := 0.09388565;
      R_f[1,0] := -0.04204104;
      R_f[1,1] := 0.43994310;
      R_f[1,2] := -0.50940818;
      R_f[1,3] := -0.20580122;
      R_f[1,4] := -0.11669060;
      R_f[1,5] := -0.12535274;
      R_f[1,6] := -0.17437693;
      R_f[1,7] := 0.09710847;
      R_f[1,8] := 0.69095361;
      R_f[1,9] := -0.05938406;
      R_f[1,10] := 0.23093407;
      R_f[1,11] := 0.13014123;
      R_f[1,12] := 0.29676151;
      R_f[1,13] := -0.05925511;
      R_f[1,14] := -0.05731449;
      R_f[1,15] := -0.06976738;
      R_f[1,16] := -0.25272533;
      R_f[1,17] := -0.25974476;
      R_f[1,18] := 0.06395108;
      R_f[1,19] := -0.02663315;
      R_f[1,20] := -0.28979155;
      R_f[1,21] := -0.76296163;
      R_f[1,22] := 1.27107012;
      R_f[1,23] := 0.14891846;
      R_f[1,24] := 0.21099623;
      R_f[1,25] := -0.11158129;
      R_f[1,26] := -0.40153420;
      R_f[1,27] := -0.29000205;
      R_f[1,28] := -0.19286913;
      R_f[1,29] := -0.01388888;
      R_f[1,30] := 0.28075165;
      R_f[1,31] := 0.47065249;
      R_f[2,0] := 0.01861088;
      R_f[2,1] := -0.03819685;
      R_f[2,2] := 0.07675387;
      R_f[2,3] := -0.08049355;
      R_f[2,4] := 0.20238465;
      R_f[2,5] := -0.63415873;
      R_f[2,6] := -0.16010195;
      R_f[2,7] := 0.20595564;
      R_f[2,8] := 0.33960930;
      R_f[2,9] := -0.38146576;
      R_f[2,10] := 0.21983975;
      R_f[2,11] := -0.28182191;
      R_f[2,12] := -0.37903464;
      R_f[2,13] := -0.32261327;
      R_f[2,14] := 0.05684026;
      R_f[2,15] := 0.11704630;
      R_f[2,16] := 0.05512832;
      R_f[2,17] := -0.31726769;
      R_f[2,18] := -0.13870730;
      R_f[2,19] := 0.15085433;
      R_f[2,20] := 0.02435878;
      R_f[2,21] := -0.60152507;
      R_f[2,22] := 0.54198354;
      R_f[2,23] := 0.02622962;
      R_f[2,24] := 0.17085208;
      R_f[2,25] := -0.24645655;
      R_f[2,26] := 0.02432794;
      R_f[2,27] := -0.42638651;
      R_f[2,28] := -0.36871403;
      R_f[2,29] := 0.21941775;
      R_f[2,30] := 0.25876975;
      R_f[2,31] := 0.23297341;
      R_f[3,0] := -0.09060316;
      R_f[3,1] := -0.12923956;
      R_f[3,2] := 0.16227835;
      R_f[3,3] := 0.20583813;
